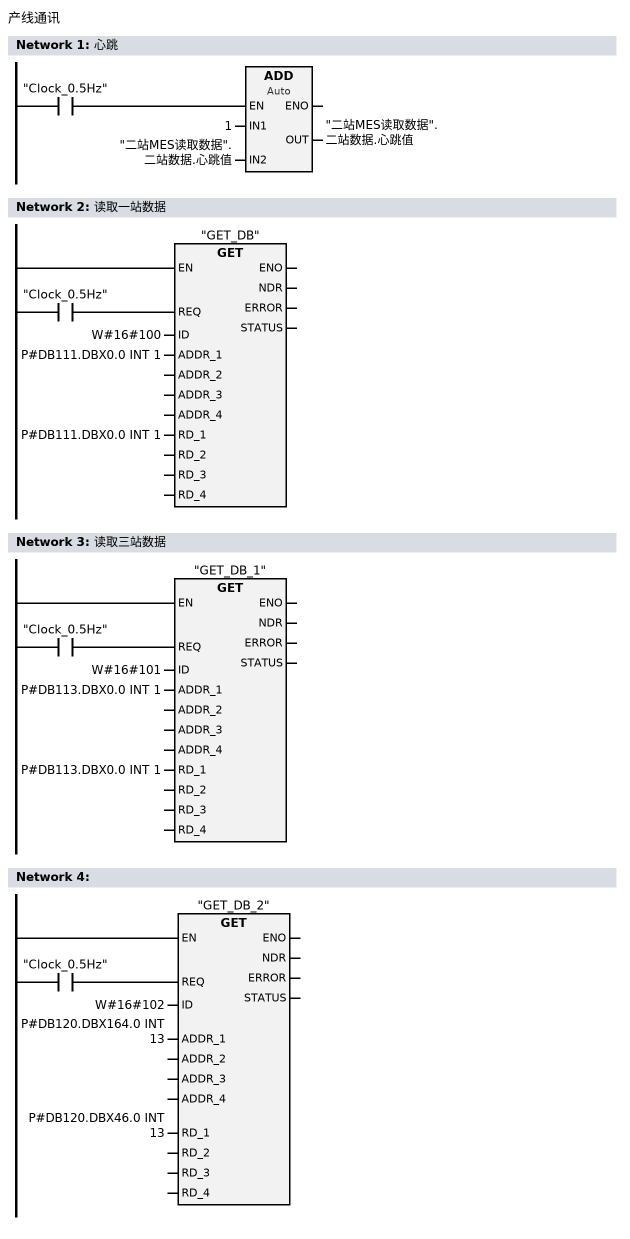
   RUNG wire#powerrail
      Contact( "Clock_0.5Hz" )
      Add(in1 := 1, in2 := "二站MES读取数据".二站数据.心跳值, out => "二站MES读取数据".二站数据.心跳值)
   END_RUNG
   // the same network as SCL:
   IF "Clock_0.5Hz" THEN "二站MES读取数据".二站数据.心跳值 := 1 + "二站MES读取数据".二站数据.心跳值; END_IF;
END_REGION

REGION Network 2: 读取一站数据
   "GET_DB"(REQ := "Clock_0.5Hz", ID := W#16#100, ADDR_1 := P#DB111.DBX0.0 INT 1, RD_1 := P#DB111.DBX0.0 INT 1);   // GET
END_REGION

REGION Network 3: 读取三站数据
   "GET_DB_1"(REQ := "Clock_0.5Hz",   // GET
              ID := W#16#101,
              ADDR_1 := P#DB113.DBX0.0 INT 1,
              RD_1 := P#DB113.DBX0.0 INT 1);
END_REGION

REGION Network 4
   "GET_DB_2"(REQ := "Clock_0.5Hz",   // GET
              ID := W#16#102,
              ADDR_1 := P#DB120.DBX164.0 INT 13,
              RD_1 := P#DB120.DBX46.0 INT 13);
END_REGION
END_FUNCTION

FUNCTION "扫码器通讯" : Void   // FC8, LAD
{ S7_Optimized_Access := 'TRUE' }
VERSION : 0.1
BEGIN

REGION Network 1
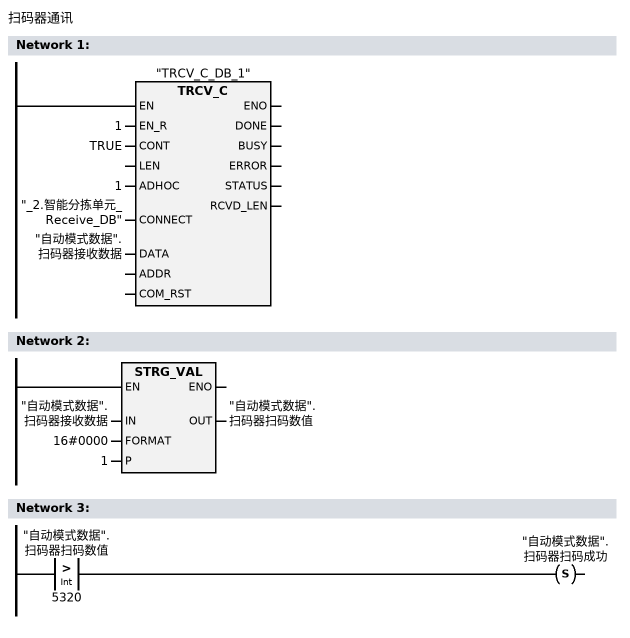
   "TRCV_C_DB_1"(EN_R := 1,   // TRCV_C
                 CONT := TRUE,
                 ADHOC := 1,
                 CONNECT := "_2.智能分拣单元_Receive_DB",
                 DATA := "自动模式数据".扫码器接收数据);
END_REGION

REGION Network 2
   STRG_VAL(IN := "自动模式数据".扫码器接收数据, FORMAT := 16#0000, P := 1, OUT => "自动模式数据".扫码器扫码数值);
END_REGION

REGION Network 3
   RUNG wire#powerrail
      { S7_Templates := "SrcType := Int" } GT_Contact(in1 := "自动模式数据".扫码器扫码数值, in2 := 5320)
      S_Coil( "自动模式数据".扫码器扫码成功 )
   END_RUNG
   // the same network as SCL:
   IF "自动模式数据".扫码器扫码数值 > 5320 THEN "自动模式数据".扫码器扫码成功 := TRUE; END_IF;
END_REGION
END_FUNCTION

FUNCTION "虚拟联动映射" : Void   // FC11, LAD
{ S7_Optimized_Access := 'TRUE' }
VERSION : 0.1
BEGIN

REGION Network 1
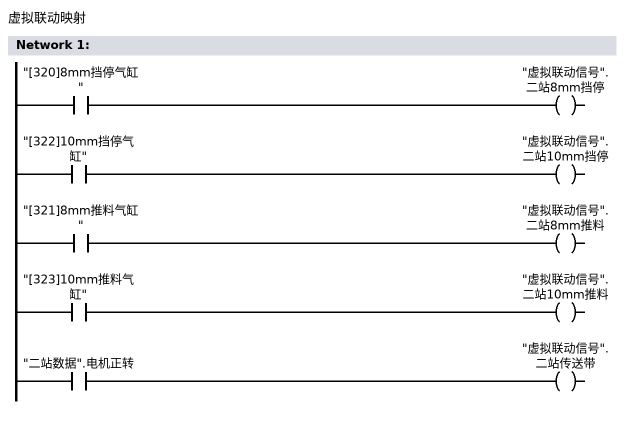
   RUNG wire#powerrail
      Contact( "[320]8mm挡停气缸" )
      Coil( "虚拟联动信号".二站8mm挡停 )
   END_RUNG
   RUNG wire#powerrail
      Contact( "[322]10mm挡停气缸" )
      Coil( "虚拟联动信号".二站10mm挡停 )
   END_RUNG
   RUNG wire#powerrail
      Contact( "[321]8mm推料气缸" )
      Coil( "虚拟联动信号".二站8mm推料 )
   END_RUNG
   RUNG wire#powerrail
      Contact( "[323]10mm推料气缸" )
      Coil( "虚拟联动信号".二站10mm推料 )
   END_RUNG
   RUNG wire#powerrail
      Contact( "二站数据".电机正转 )
      Coil( "虚拟联动信号".二站传送带 )
   END_RUNG
   // the same network as SCL:
   "虚拟联动信号".二站8mm挡停 := "[320]8mm挡停气缸";
   "虚拟联动信号".二站10mm挡停 := "[322]10mm挡停气缸";
   "虚拟联动信号".二站8mm推料 := "[321]8mm推料气缸";
   "虚拟联动信号".二站10mm推料 := "[323]10mm推料气缸";
   "虚拟联动信号".二站传送带 := "二站数据".电机正转;
END_REGION
END_FUNCTION

FUNCTION "AI视觉信号映射" : Void   // FC12, LAD
{ S7_Optimized_Access := 'TRUE' }
VERSION : 0.1
BEGIN

REGION Network 1
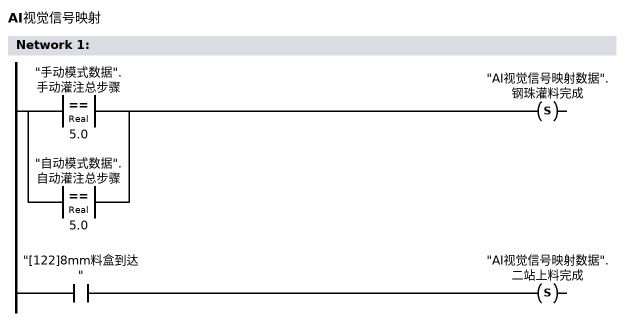
   RUNG wire#powerrail
      { S7_Templates := "SrcType := Real" } EQ_Contact(in1 := "手动模式数据".手动灌注总步骤, in2 := 5.0)
      wire#w1
      S_Coil( "AI视觉信号映射数据".钢珠灌料完成 )
   END_RUNG
   RUNG wire#powerrail
      { S7_Templates := "SrcType := Real" } EQ_Contact(in1 := "自动模式数据".自动灌注总步骤, in2 := 5.0)
   END_RUNG wire#w1
   RUNG wire#powerrail
      Contact( "[122]8mm料盒到达" )
      S_Coil( "AI视觉信号映射数据".二站上料完成 )
   END_RUNG
   // the same network as SCL:
   IF ("手动模式数据".手动灌注总步骤 = 5.0) OR ("自动模式数据".自动灌注总步骤 = 5.0) THEN "AI视觉信号映射数据".钢珠灌料完成 := TRUE; END_IF;
   IF "[122]8mm料盒到达" THEN "AI视觉信号映射数据".二站上料完成 := TRUE; END_IF;
END_REGION
END_FUNCTION

FUNCTION "MES数据映射" : Void   // FC15, LAD
{ S7_Optimized_Access := 'TRUE' }
VERSION : 0.1
BEGIN
END_FUNCTION

// ===== PLC "3.智能仓储单元"  CPU 1214C DC/DC/DC =====

VAR_GLOBAL   // PLC tag table "默认变量表"
   "System_Byte" AT %MB501 : Byte;
   "FirstScan" AT %M501.0 : Bool;
   "DiagStatusUpdate" AT %M501.1 : Bool;
   "AlwaysTRUE" AT %M501.2 : Bool;
   "AlwaysFALSE" AT %M501.3 : Bool;
   "Clock_Byte" AT %MB500 : Byte;
   "Clock_10Hz" AT %M500.0 : Bool;
   "Clock_5Hz" AT %M500.1 : Bool;
   "Clock_2.5Hz" AT %M500.2 : Bool;
   "Clock_2Hz" AT %M500.3 : Bool;
   "Clock_1.25Hz" AT %M500.4 : Bool;
   "Clock_1Hz" AT %M500.5 : Bool;
   "Clock_0.625Hz" AT %M500.6 : Bool;
   "Clock_0.5Hz" AT %M500.7 : Bool;
END_VAR

VAR_GLOBAL   // PLC tag table "第三站变量表"
   "[100]变频编码器" AT %I0.0 : Bool;
   "[101]X伺服左极限" AT %I0.1 : Bool;
   "[102]X伺服右极限" AT %I0.2 : Bool;
   "[103]X伺服原点" AT %I0.3 : Bool;
   "[104]Y伺服左极限" AT %I0.4 : Bool;
   "[105]Y伺服右极限" AT %I0.5 : Bool;
   "[106]Y原点" AT %I0.6 : Bool;
   "[107]启动" AT %I0.7 : Bool;
   "[110]停止" AT %I1.0 : Bool;
   "[111]复位" AT %I1.1 : Bool;
   "[112]急停" AT %I1.2 : Bool;
   "[113]手自动" AT %I1.3 : Bool;
   "[114]盒盖有无检测" AT %I1.4 : Bool;
   "[115]压力检测" AT %I1.5 : Bool;
   "[120]料盒到位检测" AT %I2.0 : Bool;
   "[121]不合格挡料伸出位" AT %I2.1 : Bool;
   "[122]不合格挡料缩回位" AT %I2.2 : Bool;
   "[123]滑台伸出到位" AT %I2.3 : Bool;
   "[124]滑台缩回到位" AT %I2.4 : Bool;
   "[125]]滑台左位" AT %I2.5 : Bool;
   "[126]滑台右位" AT %I2.6 : Bool;
   "[127]滑台夹爪夹紧" AT %I2.7 : Bool;
   "[130]滑台夹爪松开" AT %I3.0 : Bool;
   "[131]不合格推料伸出位" AT %I3.1 : Bool;
   "[132]不合格推料缩回位" AT %I3.2 : Bool;
   "[133]盒盖推料伸出位" AT %I3.3 : Bool;
   "[134]盒盖推料缩回位" AT %I3.4 : Bool;
   "[135]取盒盖伸出位" AT %I3.5 : Bool;
   "[136]取盒盖缩回位" AT %I3.6 : Bool;
   "[137]仓储夹爪夹紧位" AT %I3.7 : Bool;
   "[140]取盒盖上升位" AT %I4.0 : Bool;
   "[141]取盒盖下降位" AT %I4.1 : Bool;
   "[142]仓储伸出位" AT %I4.2 : Bool;
   "[143]仓储缩回位" AT %I4.3 : Bool;
   "[144]仓储上升位" AT %I4.4 : Bool;
   "[145]仓储下降位" AT %I4.5 : Bool;
   "[146]仓储夹爪松开位" AT %I4.6 : Bool;
   "[147]取料挡料伸出位" AT %I4.7 : Bool;
   "[150]取料挡料缩回位" AT %I5.0 : Bool;
   "[151]备用" AT %I5.1 : Bool;
   "[152]备用" AT %I5.2 : Bool;
   "[153]备用" AT %I5.3 : Bool;
   "轴_1_Drive_IN" AT %I68.0 : "PD_TEL3_IN";
   "轴_1_Drive_IN(1)" AT %I86.0 : "PD_TEL3_IN";
   "仓位信息" AT %IW4 : Word;
   "[303]黄色指示灯" AT %Q0.3 : Bool;
   "[304]绿色指示灯" AT %Q0.4 : Bool;
   "[305]红色指示灯" AT %Q0.5 : Bool;
   "[306]变频正转" AT %Q0.6 : Bool;
   "[307]变频反转" AT %Q0.7 : Bool;
   "[310]声光报警" AT %Q1.0 : Bool;
   "[320]不合格挡料气缸" AT %Q2.0 : Bool;
   "[321滑台伸缩气缸" AT %Q2.1 : Bool;
   "[322]滑台移动气缸" AT %Q2.2 : Bool;
   "[323]滑台夹爪气缸" AT %Q2.3 : Bool;
   "[324]不合格推料气缸" AT %Q2.4 : Bool;
   "[325]称重抬升气缸" AT %Q2.5 : Bool;
   "[326]盒盖推料气缸" AT %Q2.6 : Bool;
   "[327]取盖伸缩气缸" AT %Q2.7 : Bool;
   "[330]取盖升降气缸" AT %Q3.0 : Bool;
   "[331]取盖吸盘" AT %Q3.1 : Bool;
   "[332]仓储伸缩气缸" AT %Q3.2 : Bool;
   "[333]仓储升降气缸" AT %Q3.3 : Bool;
   "[334]仓储夹爪控制" AT %Q3.4 : Bool;
   "[335]三色灯-黄" AT %Q3.5 : Bool;
   "[336]三色灯-绿" AT %Q3.6 : Bool;
   "[337]三色灯-红" AT %Q3.7 : Bool;
   "轴_1_Drive_OUT" AT %Q64.0 : "PD_TEL3_OUT";
   "轴_1_Drive_OUT(1)" AT %Q74.0 : "PD_TEL3_OUT";
   "[154]备用4" AT %I5.4 : Bool;
   "[155]变频器故障" AT %I5.5 : Bool;
   "[156]安全光栅" AT %I5.6 : Bool;   // 1无物体2有物体
   "[157]仓位1号有无" AT %I5.7 : Bool;
   "[160]仓位2号有无" AT %I6.0 : Bool;
   "[161]仓位3号有无" AT %I6.1 : Bool;
   "[162]仓位4号有无" AT %I6.2 : Bool;
   "[163]仓位5号有无" AT %I6.3 : Bool;
   "[164]仓位6号有无" AT %I6.4 : Bool;
   "[165]仓位7号有无" AT %I6.5 : Bool;
   "[166]仓位8号有无" AT %I6.6 : Bool;
   "[167]仓位9号有无" AT %I6.7 : Bool;
   "[171]颜色检测" AT %I7.1 : Bool;
   "[170]材质检测" AT %I7.0 : Bool;
   "[311]取料挡料气缸" AT %Q1.1 : Bool;   // 滑台夹爪处挡料气缸
   "[302]备用" AT %I1.6 : Bool;
   "[301]备用" AT %I1.7 : Bool;
   "[300]备用" AT %IW108 : UInt;
   "Tag_4" AT %IW157 : Word;
   "Tag_1" AT %Q0.0 : Bool;
END_VAR

DATA_BLOCK "全局数据块"   // DB5
{ S7_Optimized_Access := 'FALSE' }
VERSION : 0.1
   VAR
      视觉检测步骤 : Real;
      称重压盖步骤 : Real;
      料盒入库步骤 : Real;
      仓储总步骤 : Real;
      重量存储库 : Struct
         "1" : Int;
         "2" : Int;
         "3" : Int;
         "4" : Int;
         "5" : Int;
         "6" : Int;
         "7" : Int;
         "8" : Int;
      END_STRUCT;
      变频器启动 : Bool;
      入站扫码数据 : String[16];
      入站扫码数值 : Int;
      入站扫码成功 : Bool;
      入库扫码数据 : String[16];
      入库扫码数值 : Int;
      入库扫码成功 : Bool;
      视觉检测等待时间 : Time := T#2S;
      不合格产品计数 : Int;
      合格产品计数 : Int;
      上个完成订单ID : Int;
      手动模式步骤 : Real;
      手动存储仓位 : Int := 5;
   END_VAR
BEGIN
END_DATA_BLOCK

DATA_BLOCK "初始化数据"   // DB8
{ S7_Optimized_Access := 'FALSE' }
VERSION : 0.1
   VAR
      手动模式 : Bool;
      自动模式 : Bool;
      自动运行模式 : Bool;
      初始化步骤 : Int;
      初始化完成 : Bool;
      初始化中 : Bool;
      初始化故障 : Bool;
      急停状态 : Bool;
      安全光栅被挡 : Bool;
      黄灯_内部 : Bool;
      红灯_内部 : Bool;
      绿灯_内部 : Bool;
      报警等级 : Int;
      报警确认按钮 : Bool;
      报警总输出 : Bool;
   END_VAR
BEGIN
END_DATA_BLOCK

DATA_BLOCK "状态控制数据"   // DB44
{ S7_Optimized_Access := 'FALSE' }
VERSION : 0.1
   VAR
      在线状态 : Bool;   // PLC已经上电
      忙碌状态 : Bool;   // 三站已经接单
      空闲状态 : Bool;   // 三站准备就绪(没急停，初始化已经完成，光栅没被挡)
      故障状态 : Bool;   // 报警、光栅被挡
   END_VAR
BEGIN
END_DATA_BLOCK

DATA_BLOCK "三站MES读取数据"   // DB120
{ S7_Optimized_Access := 'FALSE' }
VERSION : 0.1
   VAR
      三站数据 : Struct
         在线状态 : Int;
         运行模式 : Int;   // 0 手动 / 1 自动待机 / 2 自动运行
         忙碌状态 : Int;   // 0 空闲 / 1 忙碌
         故障状态 : Int;   // 0 = 无故障
         当前订单ID : Int;   // 当前处理的订单
         当前步骤 : Real;
         心跳值 : Int;
         三站完成 : Bool;
         保留 : Bool;
         保留_1 : Bool;
         保留_2 : Bool;
         保留_3 : Bool;
         保留_4 : Bool;
         保留_5 : Bool;
         保留_6 : Bool;
         仓位状态 : Array[0..8] of Bool;
         入站扫码数据 : Int;
         入库扫码数据 : Int;
         称重数据 : Int;
         产品合格状态 : Int;
         合格产品计数 : Int;
         不合格产品计数 : Int;
         X轴当前位置 : Real;
         Y轴当前位置 : Real;
         完成订单ID : Int;
         三站保留数据 : Array[0..8] of Int;
      END_STRUCT;
      订单数据 : Struct
         订单id : Int;
         ab物料 : Int;   // 1A，2B，3不需要
         小钢珠数量 : Int;
         大钢珠数量 : Int;
         存储仓位 : Int;
         当前订单完成 : Bool;
         开始信号 : Int;
         复位信号 : Int;
         订单保留数据 : Array[0..4] of Int;
      END_STRUCT;
   END_VAR
BEGIN
END_DATA_BLOCK

// folder: System blocks/Program resources

DATA_BLOCK "IEC_Timer_0_DB_7"   // DB7
{ S7_Optimized_Access := 'TRUE' }
AUTHOR : Simatic
FAMILY : IEC
NAME : IEC_TMR
VERSION : 1.0
// stored: InstanceOfName IEC_TIMER
"IEC_TIMER"
BEGIN
END_DATA_BLOCK

DATA_BLOCK "IEC_Timer_0_DB_4"   // DB9
{ S7_Optimized_Access := 'TRUE' }
AUTHOR : Simatic
FAMILY : IEC
NAME : IEC_TMR
VERSION : 1.0
// stored: InstanceOfName IEC_TIMER
"IEC_TIMER"
BEGIN
END_DATA_BLOCK

DATA_BLOCK "IEC_Timer_0_DB"   // DB13
{ S7_Optimized_Access := 'TRUE' }
AUTHOR : Simatic
FAMILY : IEC
NAME : IEC_TMR
VERSION : 1.0
// stored: InstanceOfName IEC_TIMER
"IEC_TIMER"
BEGIN
END_DATA_BLOCK

DATA_BLOCK "IEC_Timer_0_DB_1"   // DB14
{ S7_Optimized_Access := 'TRUE' }
AUTHOR : Simatic
FAMILY : IEC
NAME : IEC_TMR
VERSION : 1.0
// stored: InstanceOfName IEC_TIMER
"IEC_TIMER"
BEGIN
END_DATA_BLOCK

DATA_BLOCK "IEC_Timer_0_DB_2"   // DB15
{ S7_Optimized_Access := 'TRUE' }
AUTHOR : Simatic
FAMILY : IEC
NAME : IEC_TMR
VERSION : 1.0
// stored: InstanceOfName IEC_TIMER
"IEC_TIMER"
BEGIN
END_DATA_BLOCK

DATA_BLOCK "IEC_Timer_0_DB_3"   // DB16
{ S7_Optimized_Access := 'TRUE' }
AUTHOR : Simatic
FAMILY : IEC
NAME : IEC_TMR
VERSION : 1.0
// stored: InstanceOfName IEC_TIMER
"IEC_TIMER"
BEGIN
END_DATA_BLOCK

DATA_BLOCK "IEC_Timer_0_DB_5"   // DB18
{ S7_Optimized_Access := 'TRUE' }
AUTHOR : Simatic
FAMILY : IEC
NAME : IEC_TMR
VERSION : 1.0
// stored: InstanceOfName IEC_TIMER
"IEC_TIMER"
BEGIN
END_DATA_BLOCK

DATA_BLOCK "IEC_Timer_0_DB_6"   // DB19
{ S7_Optimized_Access := 'TRUE' }
AUTHOR : Simatic
FAMILY : IEC
NAME : IEC_TMR
VERSION : 1.0
// stored: InstanceOfName IEC_TIMER
"IEC_TIMER"
BEGIN
END_DATA_BLOCK

DATA_BLOCK "IEC_Timer_0_DB_8"   // DB28
{ S7_Optimized_Access := 'TRUE' }
AUTHOR : Simatic
FAMILY : IEC
NAME : IEC_TMR
VERSION : 1.0
// stored: InstanceOfName IEC_TIMER
"IEC_TIMER"
BEGIN
END_DATA_BLOCK

DATA_BLOCK "IEC_Timer_0_DB_9"   // DB29
{ S7_Optimized_Access := 'TRUE' }
AUTHOR : Simatic
FAMILY : IEC
NAME : IEC_TMR
VERSION : 1.0
// stored: InstanceOfName IEC_TIMER
"IEC_TIMER"
BEGIN
END_DATA_BLOCK

DATA_BLOCK "IEC_Timer_0_DB_10"   // DB30
{ S7_Optimized_Access := 'TRUE' }
AUTHOR : Simatic
FAMILY : IEC
NAME : IEC_TMR
VERSION : 1.0
// stored: InstanceOfName IEC_TIMER
"IEC_TIMER"
BEGIN
END_DATA_BLOCK

DATA_BLOCK "IEC_Timer_0_DB_11"   // DB31
{ S7_Optimized_Access := 'TRUE' }
AUTHOR : Simatic
FAMILY : IEC
NAME : IEC_TMR
VERSION : 1.0
// stored: InstanceOfName IEC_TIMER
"IEC_TIMER"
BEGIN
END_DATA_BLOCK

DATA_BLOCK "IEC_Timer_0_DB_12"   // DB32
{ S7_Optimized_Access := 'TRUE' }
AUTHOR : Simatic
FAMILY : IEC
NAME : IEC_TMR
VERSION : 1.0
// stored: InstanceOfName IEC_TIMER
"IEC_TIMER"
BEGIN
END_DATA_BLOCK

DATA_BLOCK "IEC_Timer_0_DB_13"   // DB33
{ S7_Optimized_Access := 'TRUE' }
AUTHOR : Simatic
FAMILY : IEC
NAME : IEC_TMR
VERSION : 1.0
// stored: InstanceOfName IEC_TIMER
"IEC_TIMER"
BEGIN
END_DATA_BLOCK

DATA_BLOCK "_3.智能仓储单元_Receive_DB"   // DB35
{ S7_Optimized_Access := 'TRUE' }
AUTHOR : SIMATIC
FAMILY : MC7Plus
NAME : TC_IP_v4
VERSION : 1.0
// stored: InstanceOfName TCON_IP_v4
"TCON_IP_v4"
BEGIN
   ID := 104;
   InterfaceId := 64;
   LocalPort := 8899;
   RemotePort := 8899;
   RemoteAddress.ADDR[1] := 192;
   RemoteAddress.ADDR[2] := 168;
   RemoteAddress.ADDR[3] := 40;
   RemoteAddress.ADDR[4] := 103;
END_DATA_BLOCK

DATA_BLOCK "IEC_Timer_0_DB_17"   // DB37
{ S7_Optimized_Access := 'TRUE' }
AUTHOR : Simatic
FAMILY : IEC
NAME : IEC_TMR
VERSION : 1.0
// stored: InstanceOfName IEC_TIMER
"IEC_TIMER"
BEGIN
END_DATA_BLOCK

DATA_BLOCK "IEC_Timer_0_DB_18"   // DB38
{ S7_Optimized_Access := 'TRUE' }
AUTHOR : Simatic
FAMILY : IEC
NAME : IEC_TMR
VERSION : 1.0
// stored: InstanceOfName IEC_TIMER
"IEC_TIMER"
BEGIN
END_DATA_BLOCK

DATA_BLOCK "IEC_Timer_0_DB_19"   // DB39
{ S7_Optimized_Access := 'TRUE' }
AUTHOR : Simatic
FAMILY : IEC
NAME : IEC_TMR
VERSION : 1.0
// stored: InstanceOfName IEC_TIMER
"IEC_TIMER"
BEGIN
END_DATA_BLOCK

DATA_BLOCK "IEC_Timer_0_DB_16"   // DB40
{ S7_Optimized_Access := 'TRUE' }
AUTHOR : Simatic
FAMILY : IEC
NAME : IEC_TMR
VERSION : 1.0
// stored: InstanceOfName IEC_TIMER
"IEC_TIMER"
BEGIN
END_DATA_BLOCK

DATA_BLOCK "_3.智能仓储单元_Receive_DB_1"   // DB41
{ S7_Optimized_Access := 'TRUE' }
AUTHOR : SIMATIC
FAMILY : MC7Plus
NAME : TC_IP_v4
VERSION : 1.0
// stored: InstanceOfName TCON_IP_v4
"TCON_IP_v4"
BEGIN
   ID := 107;
   InterfaceId := 64;
   LocalPort := 8899;
   RemotePort := 8899;
   RemoteAddress.ADDR[1] := 192;
   RemoteAddress.ADDR[2] := 168;
   RemoteAddress.ADDR[3] := 40;
   RemoteAddress.ADDR[4] := 102;
END_DATA_BLOCK

DATA_BLOCK "IEC_Timer_0_DB_20"   // DB42
{ S7_Optimized_Access := 'TRUE' }
AUTHOR : Simatic
FAMILY : IEC
NAME : IEC_TMR
VERSION : 1.0
// stored: InstanceOfName IEC_TIMER
"IEC_TIMER"
BEGIN
END_DATA_BLOCK

DATA_BLOCK "IEC_Timer_0_DB_14"   // DB45
{ S7_Optimized_Access := 'TRUE' }
AUTHOR : Simatic
FAMILY : IEC
NAME : IEC_TMR
VERSION : 1.0
// stored: InstanceOfName IEC_TIMER
"IEC_TIMER"
BEGIN
END_DATA_BLOCK

DATA_BLOCK "IEC_Timer_0_DB_15"   // DB46
{ S7_Optimized_Access := 'TRUE' }
AUTHOR : Simatic
FAMILY : IEC
NAME : IEC_TMR
VERSION : 1.0
// stored: InstanceOfName IEC_TIMER
"IEC_TIMER"
BEGIN
END_DATA_BLOCK

DATA_BLOCK "IEC_Timer_0_DB_21"   // DB47
{ S7_Optimized_Access := 'TRUE' }
AUTHOR : Simatic
FAMILY : IEC
NAME : IEC_TMR
VERSION : 1.0
// stored: InstanceOfName IEC_TIMER
"IEC_TIMER"
BEGIN
END_DATA_BLOCK

DATA_BLOCK "IEC_Timer_0_DB_22"   // DB48
{ S7_Optimized_Access := 'TRUE' }
AUTHOR : Simatic
FAMILY : IEC
NAME : IEC_TMR
VERSION : 1.0
// stored: InstanceOfName IEC_TIMER
"IEC_TIMER"
BEGIN
END_DATA_BLOCK

DATA_BLOCK "IEC_Timer_0_DB_23"   // DB49
{ S7_Optimized_Access := 'TRUE' }
AUTHOR : Simatic
FAMILY : IEC
NAME : IEC_TMR
VERSION : 1.0
// stored: InstanceOfName IEC_TIMER
"IEC_TIMER"
BEGIN
END_DATA_BLOCK

DATA_BLOCK "IEC_Timer_0_DB_24"   // DB50
{ S7_Optimized_Access := 'TRUE' }
AUTHOR : Simatic
FAMILY : IEC
NAME : IEC_TMR
VERSION : 1.0
// stored: InstanceOfName IEC_TIMER
"IEC_TIMER"
BEGIN
END_DATA_BLOCK

DATA_BLOCK "IEC_Timer_0_DB_25"   // DB51
{ S7_Optimized_Access := 'TRUE' }
AUTHOR : Simatic
FAMILY : IEC
NAME : IEC_TMR
VERSION : 1.0
// stored: InstanceOfName IEC_TIMER
"IEC_TIMER"
BEGIN
END_DATA_BLOCK

DATA_BLOCK "IEC_Timer_0_DB_26"   // DB52
{ S7_Optimized_Access := 'TRUE' }
AUTHOR : Simatic
FAMILY : IEC
NAME : IEC_TMR
VERSION : 1.0
// stored: InstanceOfName IEC_TIMER
"IEC_TIMER"
BEGIN
END_DATA_BLOCK

DATA_BLOCK "IEC_Timer_0_DB_27"   // DB53
{ S7_Optimized_Access := 'TRUE' }
AUTHOR : Simatic
FAMILY : IEC
NAME : IEC_TMR
VERSION : 1.0
// stored: InstanceOfName IEC_TIMER
"IEC_TIMER"
BEGIN
END_DATA_BLOCK

DATA_BLOCK "IEC_Timer_0_DB_28"   // DB54
{ S7_Optimized_Access := 'TRUE' }
AUTHOR : Simatic
FAMILY : IEC
NAME : IEC_TMR
VERSION : 1.0
// stored: InstanceOfName IEC_TIMER
"IEC_TIMER"
BEGIN
END_DATA_BLOCK

DATA_BLOCK "IEC_Timer_0_DB_29"   // DB55
{ S7_Optimized_Access := 'TRUE' }
AUTHOR : Simatic
FAMILY : IEC
NAME : IEC_TMR
VERSION : 1.0
// stored: InstanceOfName IEC_TIMER
"IEC_TIMER"
BEGIN
END_DATA_BLOCK

DATA_BLOCK "IEC_Timer_0_DB_30"   // DB56
{ S7_Optimized_Access := 'TRUE' }
AUTHOR : Simatic
FAMILY : IEC
NAME : IEC_TMR
VERSION : 1.0
// stored: InstanceOfName IEC_TIMER
"IEC_TIMER"
BEGIN
END_DATA_BLOCK

DATA_BLOCK "IEC_Timer_0_DB_31"   // DB57
{ S7_Optimized_Access := 'TRUE' }
AUTHOR : Simatic
FAMILY : IEC
NAME : IEC_TMR
VERSION : 1.0
// stored: InstanceOfName IEC_TIMER
"IEC_TIMER"
BEGIN
END_DATA_BLOCK

DATA_BLOCK "IEC_Timer_0_DB_32"   // DB58
{ S7_Optimized_Access := 'TRUE' }
AUTHOR : Simatic
FAMILY : IEC
NAME : IEC_TMR
VERSION : 1.0
// stored: InstanceOfName IEC_TIMER
"IEC_TIMER"
BEGIN
END_DATA_BLOCK

DATA_BLOCK "IEC_Timer_0_DB_33"   // DB59
{ S7_Optimized_Access := 'TRUE' }
AUTHOR : Simatic
FAMILY : IEC
NAME : IEC_TMR
VERSION : 1.0
// stored: InstanceOfName IEC_TIMER
"IEC_TIMER"
BEGIN
END_DATA_BLOCK

DATA_BLOCK "IEC_Timer_0_DB_34"   // DB60
{ S7_Optimized_Access := 'TRUE' }
AUTHOR : Simatic
FAMILY : IEC
NAME : IEC_TMR
VERSION : 1.0
// stored: InstanceOfName IEC_TIMER
"IEC_TIMER"
BEGIN
END_DATA_BLOCK

DATA_BLOCK "IEC_Timer_0_DB_35"   // DB61
{ S7_Optimized_Access := 'TRUE' }
AUTHOR : Simatic
FAMILY : IEC
NAME : IEC_TMR
VERSION : 1.0
// stored: InstanceOfName IEC_TIMER
"IEC_TIMER"
BEGIN
END_DATA_BLOCK

// folder: 运动控制

DATA_BLOCK "运动控制数据2"   // DB1
{ S7_Optimized_Access := 'FALSE' }
VERSION : 0.1
   VAR
      X轴位置 : Real;
      Y轴位置 : Real;
      称重抓取x值 : Real := -82.0;
      称重抓取y值 : Real := 537.0;
      扫码位x值 : Real := -29.0;
      扫码位y值 : Real := 382.0;
      abc位x值 : Real := 151.0;
      def位x值 : Real := -32.0;
      ghi位x值 : Real := -208.0;
      adg位y值 : Real := -231.0;
      bef位y值 : Real := -51.0;
      cfi位y值 : Real := 121.0;
      "出仓位x值-420.38" : Real := -416.0;
      "出仓位y值162.88" : Real := 152.0;
      X值统一入库位 : Bool;
      Y值统一入库位 : Bool;
      X值计算 : Int;
      Y值计算 : Int;
      Y值转换后 : Int;
   END_VAR
BEGIN
END_DATA_BLOCK

DATA_BLOCK "运动控制数据1"   // DB43
{ S7_Optimized_Access := 'FALSE' }
VERSION : 0.1
   VAR
      轴初始化按钮 : Bool;
      轴初始化完成 : Bool;
      轴初始化步骤 : Int;
      轴初始化错误 : Bool;
      X轴机械手错误输出 : Bool;
      Y轴机械手错误输出 : Bool;
      X轴使能按钮 : Bool;
      X轴使能状态 : Bool;
      X轴使能错误 : Bool;
      X轴复位按钮 : Bool;
      X轴复位完成 : Bool;
      X轴复位错误 : Bool;
      X轴回原位按钮 : Bool;
      X轴回原位完成 : Bool;
      X轴回原位错误 : Bool;
      X轴绝对定位按钮 : Bool;
      X轴绝对定位完成 : Bool;
      X轴绝对定位错误 : Bool;
      Y轴使能按钮 : Bool;
      Y轴使能状态 : Bool;
      Y轴使能错误 : Bool;
      Y轴复位按钮 : Bool;
      Y轴复位完成 : Bool;
      Y轴复位错误 : Bool;
      Y轴回原位按钮 : Bool;
      Y轴回原位完成 : Bool;
      Y轴回原位错误 : Bool;
      Y轴绝对定位按钮 : Bool;
      Y轴绝对定位完成 : Bool;
      Y轴绝对定位错误 : Bool;
   END_VAR
BEGIN
END_DATA_BLOCK

// folder: 通讯模块

DATA_BLOCK "虚实联动信号"   // DB4
{ S7_Optimized_Access := 'FALSE' }
VERSION : 0.1
   VAR
      变频正转 : Bool;
      变频反转 : Bool;
      滑台移动气缸 : Bool;
      滑台伸缩气缸 : Bool;
      仓储伸缩气缸 : Bool;
      仓储升降气缸 : Bool;
      称重抬升气缸 : Bool;
      不合格推料气缸 : Bool;
      不合格挡料气缸 : Bool;
      取料挡料气缸 : Bool;
      取盖伸缩气缸 : Bool;
      取盖升降气缸 : Bool;
      盒盖推料气缸 : Bool;
      滑台夹爪气缸 : Bool;
      仓储夹爪控制 : Bool;
      取盖吸盘 : Bool;
   END_VAR
BEGIN
END_DATA_BLOCK

DATA_BLOCK "称重数据"   // DB12
{ S7_Optimized_Access := 'FALSE' }
VERSION : 0.1
   VAR
      称重 : Struct
         称重数据 : Int;
         称重数据接收 : Int;
      END_STRUCT;
   END_VAR
BEGIN
END_DATA_BLOCK

DATA_BLOCK "一站数据"   // DB111
{ S7_Optimized_Access := 'FALSE' }
VERSION : 0.1
   VAR
      一站完成 : Bool;
      复位完成 : Bool;
      一站就绪 : Bool;
      一站忙碌 : Bool;
      一站请求二站接收 : Bool;
      一站可接单 : Bool;
      数据7 : Bool;
      数据8 : Bool;
      数据9 : Bool;
      数据10 : Bool;
      数据11 : Bool;
      数据12 : Bool;
      数据13 : Bool;
      数据14 : Bool;
   END_VAR
BEGIN
END_DATA_BLOCK

DATA_BLOCK "二站数据"   // DB112
{ S7_Optimized_Access := 'FALSE' }
VERSION : 0.1
   VAR
      二站完成 : Bool;
      二站已接收 : Bool;
      复位完成 : Bool;
      空闲状态 : Bool;
      电机正转 : Bool;
      二站忙碌 : Bool;
      二站请求三站接收 : Bool;
      二站可接收 : Bool;
      数据17 : Bool;
      数据18 : Bool;
      数据19 : Bool;
      数据20 : Bool;
      数据21 : Bool;
   END_VAR
BEGIN
END_DATA_BLOCK

DATA_BLOCK "三站数据"   // DB113
{ S7_Optimized_Access := 'FALSE' }
VERSION : 0.1
   VAR
      三站完成 : Bool;
      三站已接收 : Bool;
      复位完成 : Bool;
      空闲状态 : Bool;
      出现废料 : Bool;
      安全光栅 : Bool;
      三站可接收 : Bool;
      三站忙碌 : Bool;
      数据23 : Bool;
      数据24 : Bool;
      数据25 : Bool;
      数据26 : Bool;
      数据27 : Bool;
      数据28 : Bool;
      数据29 : Bool;
   END_VAR
BEGIN
END_DATA_BLOCK

DATA_BLOCK "AI视觉信号映射数据"   // DB116
{ S7_Optimized_Access := 'TRUE' }
VERSION : 0.1
   VAR
      三站压盖完成 : Bool;
      三站入库完成 : Bool;
   END_VAR
BEGIN
END_DATA_BLOCK

// folder: (top level)

DATA_BLOCK "X轴机械手"   // DB2, Motion_DB
{ S7_Optimized_Access := 'TRUE' }
AUTHOR : SIMATIC
FAMILY : BasicMC
NAME : TO_PosAx
VERSION : 7.0
// stored: InstanceOfName TO_PositioningAxis
"TO_PositioningAxis"
BEGIN
   // Axis.HomingReferencePointSwitch_AddressCU = %I0.3
   // Axis.PositionLimitsMax_AddressCU = %I0.1
   // Axis.PositionLimitsMin_AddressCU = %I0.2
   // Axis.Encoder.TelegramAddressOutCU = %Q74.0
   // Axis.Encoder.TelegramAddressInCU = %I86.0
   // Axis.Encoder.DoNameCU = SINAMICS-V90-PN_2.驱动_1_编码器1
   // Axis.Drive.TelegramAddressOutCU = %Q74.0
   // Axis.Drive.TelegramAddressInCU = %I86.0
   // Axis.Drive.TelegramType = 2
   // Axis.Drive.DoNameCU = SINAMICS-V90-PN_2.驱动_1
   // Axis.LengthUnitNormalized.Distance = 1013
   // Axis.Encoder.SelectedHscIndexCU = -1
   // Axis.Encoder.DbTypeCU = Classic
   // Axis.Drive.DbTypeCU = Classic
END_DATA_BLOCK

DATA_BLOCK "Y轴机械手"   // DB3, Motion_DB
{ S7_Optimized_Access := 'TRUE' }
AUTHOR : SIMATIC
FAMILY : BasicMC
NAME : TO_PosAx
VERSION : 7.0
// stored: InstanceOfName TO_PositioningAxis
"TO_PositioningAxis"
BEGIN
   // Axis.HomingReferencePointSwitch_AddressCU = %I0.6
   // Axis.PositionLimitsMax_AddressCU = %I0.4
   // Axis.PositionLimitsMin_AddressCU = %I0.5
   // Axis.Encoder.TelegramAddressOutCU = %Q64.0
   // Axis.Encoder.TelegramAddressInCU = %I68.0
   // Axis.Encoder.DoNameCU = SINAMICS-V90-PN_1.驱动_1_编码器1
   // Axis.Drive.TelegramAddressOutCU = %Q64.0
   // Axis.Drive.TelegramAddressInCU = %I68.0
   // Axis.Drive.TelegramType = 2
   // Axis.Drive.DoNameCU = SINAMICS-V90-PN_1.驱动_1
   // Axis.LengthUnitNormalized.Distance = 1013
   // Axis.Encoder.SelectedHscIndexCU = -1
   // Axis.Encoder.DbTypeCU = Classic
   // Axis.Drive.DbTypeCU = Classic
END_DATA_BLOCK

FUNCTION "0.初始化" : Void   // FC5, LAD
{ S7_Optimized_Access := 'TRUE' }
VERSION : 0.1
   VAR_TEMP   // added for the SCL form of the ladder/FBD networks
      _w1 : Bool;
      _w2 : Bool;
   END_VAR
BEGIN

REGION Network 1: 模式切换
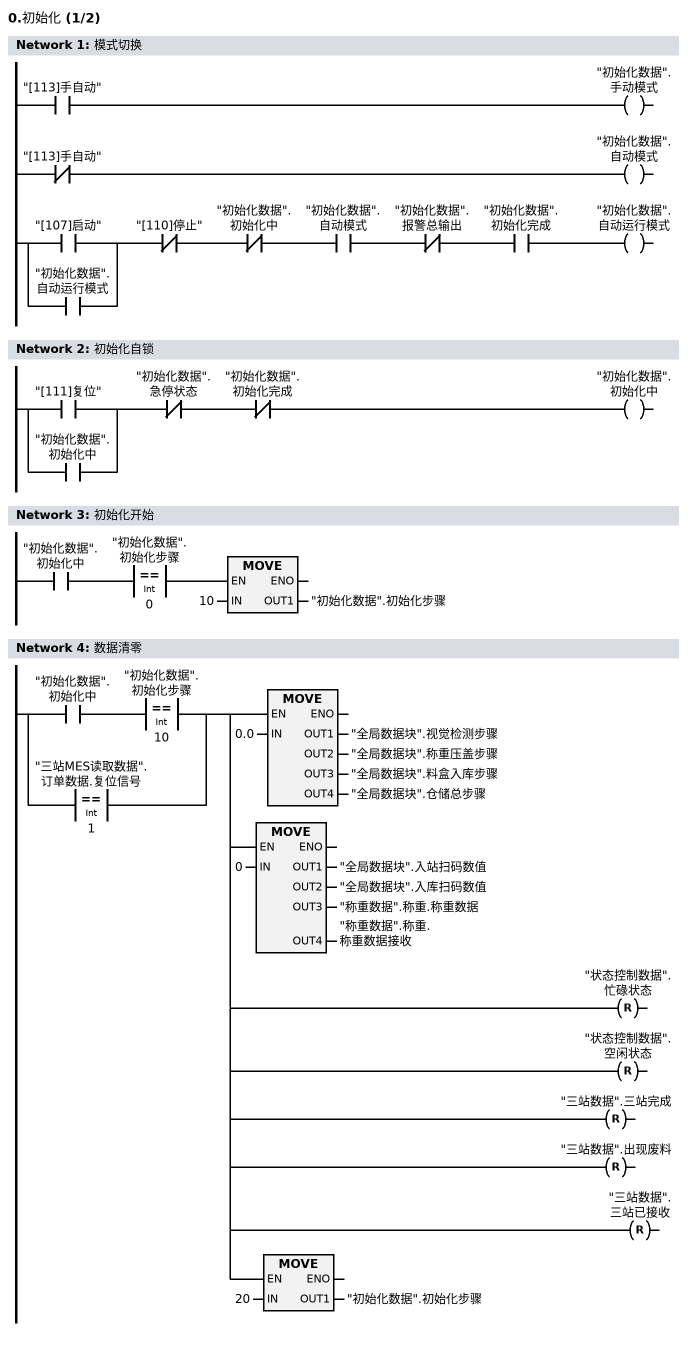
   RUNG wire#powerrail
      Contact( "[113]手自动" )
      Coil( "初始化数据".手动模式 )
   END_RUNG
   RUNG wire#powerrail
      I_Contact( "[113]手自动" )
      Coil( "初始化数据".自动模式 )
   END_RUNG
   RUNG wire#powerrail
      Contact( "[107]启动" )
      wire#w1
      I_Contact( "[110]停止" )
      I_Contact( "初始化数据".初始化中 )
      Contact( "初始化数据".自动模式 )
      I_Contact( "初始化数据".报警总输出 )
      Contact( "初始化数据".初始化完成 )
      Coil( "初始化数据".自动运行模式 )
   END_RUNG
   RUNG wire#powerrail
      Contact( "初始化数据".自动运行模式 )
   END_RUNG wire#w1
   // the same network as SCL:
   "初始化数据".手动模式 := "[113]手自动";
   "初始化数据".自动模式 := NOT "[113]手自动";
   "初始化数据".自动运行模式 := ("[107]启动" OR "初始化数据".自动运行模式) AND NOT "[110]停止" AND NOT "初始化数据".初始化中 AND "初始化数据".自动模式 AND NOT "初始化数据".报警总输出 AND "初始化数据".初始化完成;
END_REGION

REGION Network 2: 初始化自锁
   RUNG wire#powerrail
      Contact( "[111]复位" )
      wire#w1
      I_Contact( "初始化数据".急停状态 )
      I_Contact( "初始化数据".初始化完成 )
      Coil( "初始化数据".初始化中 )
   END_RUNG
   RUNG wire#powerrail
      Contact( "初始化数据".初始化中 )
   END_RUNG wire#w1
   // the same network as SCL:
   "初始化数据".初始化中 := ("[111]复位" OR "初始化数据".初始化中) AND NOT "初始化数据".急停状态 AND NOT "初始化数据".初始化完成;
END_REGION

REGION Network 3: 初始化开始
   RUNG wire#powerrail
      Contact( "初始化数据".初始化中 )
      { S7_Templates := "SrcType := Int" } EQ_Contact(in1 := "初始化数据".初始化步骤, in2 := 0)
      Move(in := 10, out1 => "初始化数据".初始化步骤)
   END_RUNG
   // the same network as SCL:
   IF "初始化数据".初始化中 AND ("初始化数据".初始化步骤 = 0) THEN "初始化数据".初始化步骤 := 10; END_IF;
END_REGION

REGION Network 4: 数据清零
   RUNG wire#powerrail
      Contact( "初始化数据".初始化中 )
      { S7_Templates := "SrcType := Int" } EQ_Contact(in1 := "初始化数据".初始化步骤, in2 := 10)
      wire#w1
      Move(in := 0.0, out1 => "全局数据块".视觉检测步骤, out2 => "全局数据块".称重压盖步骤, out3 => "全局数据块".料盒入库步骤, out4 => "全局数据块".仓储总步骤)
   END_RUNG
   RUNG wire#powerrail
      { S7_Templates := "SrcType := Int" } EQ_Contact(in1 := "三站MES读取数据".订单数据.复位信号, in2 := 1)
   END_RUNG wire#w1
   RUNG wire#w1
      Move(in := 0, out1 => "全局数据块".入站扫码数值, out2 => "全局数据块".入库扫码数值, out3 => "称重数据".称重.称重数据, out4 => "称重数据".称重.称重数据接收)
   END_RUNG
   RUNG wire#w1
      R_Coil( "状态控制数据".忙碌状态 )
   END_RUNG
   RUNG wire#w1
      R_Coil( "状态控制数据".空闲状态 )
   END_RUNG
   RUNG wire#w1
      R_Coil( "三站数据".三站完成 )
   END_RUNG
   RUNG wire#w1
      R_Coil( "三站数据".出现废料 )
   END_RUNG
   RUNG wire#w1
      R_Coil( "三站数据".三站已接收 )
   END_RUNG
   RUNG wire#w1
      Move(in := 20, out1 => "初始化数据".初始化步骤)
   END_RUNG
   // the same network as SCL:
   IF ("初始化数据".初始化中 AND ("初始化数据".初始化步骤 = 10)) OR ("三站MES读取数据".订单数据.复位信号 = 1) THEN
       "全局数据块".视觉检测步骤 := 0.0;
       "全局数据块".称重压盖步骤 := 0.0;
       "全局数据块".料盒入库步骤 := 0.0;
       "全局数据块".仓储总步骤 := 0.0;
       "全局数据块".入站扫码数值 := 0;
       "全局数据块".入库扫码数值 := 0;
       "称重数据".称重.称重数据 := 0;
       "称重数据".称重.称重数据接收 := 0;
       "状态控制数据".忙碌状态 := FALSE;
       "状态控制数据".空闲状态 := FALSE;
       "三站数据".三站完成 := FALSE;
       "三站数据".出现废料 := FALSE;
       "三站数据".三站已接收 := FALSE;
       "初始化数据".初始化步骤 := 20;
   END_IF;
END_REGION

REGION Network 6: 气缸复位
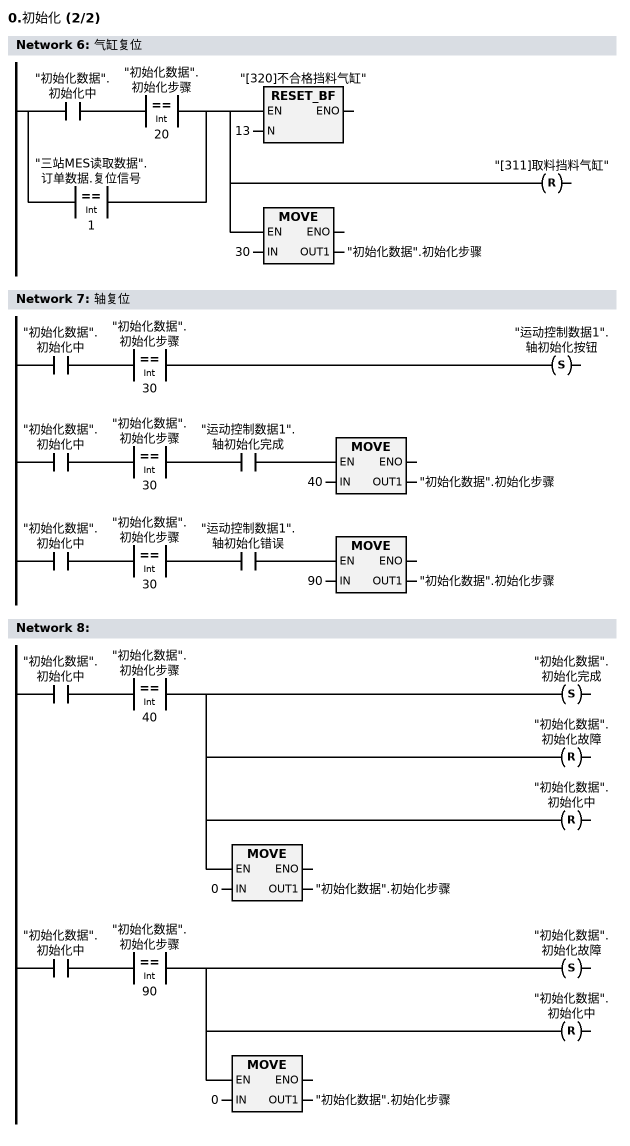
   // no SCL statement known for RBitfield: written as a call
   #_w1 := ("初始化数据".初始化中 AND ("初始化数据".初始化步骤 = 20)) OR ("三站MES读取数据".订单数据.复位信号 = 1);
   IF #_w1 THEN
       RESET_BF(operand := "[320]不合格挡料气缸", n := 13);
       "[311]取料挡料气缸" := FALSE;
       "初始化数据".初始化步骤 := 30;
   END_IF;
END_REGION

REGION Network 7: 轴复位
   RUNG wire#powerrail
      Contact( "初始化数据".初始化中 )
      { S7_Templates := "SrcType := Int" } EQ_Contact(in1 := "初始化数据".初始化步骤, in2 := 30)
      S_Coil( "运动控制数据1".轴初始化按钮 )
   END_RUNG
   RUNG wire#powerrail
      Contact( "初始化数据".初始化中 )
      { S7_Templates := "SrcType := Int" } EQ_Contact(in1 := "初始化数据".初始化步骤, in2 := 30)
      Contact( "运动控制数据1".轴初始化完成 )
      Move(in := 40, out1 => "初始化数据".初始化步骤)
   END_RUNG
   RUNG wire#powerrail
      Contact( "初始化数据".初始化中 )
      { S7_Templates := "SrcType := Int" } EQ_Contact(in1 := "初始化数据".初始化步骤, in2 := 30)
      Contact( "运动控制数据1".轴初始化错误 )
      Move(in := 90, out1 => "初始化数据".初始化步骤)
   END_RUNG
   // the same network as SCL:
   IF "初始化数据".初始化中 AND ("初始化数据".初始化步骤 = 30) THEN "运动控制数据1".轴初始化按钮 := TRUE; END_IF;
   IF "初始化数据".初始化中 AND ("初始化数据".初始化步骤 = 30) AND "运动控制数据1".轴初始化完成 THEN "初始化数据".初始化步骤 := 40; END_IF;
   IF "初始化数据".初始化中 AND ("初始化数据".初始化步骤 = 30) AND "运动控制数据1".轴初始化错误 THEN "初始化数据".初始化步骤 := 90; END_IF;
END_REGION

REGION Network 8
   RUNG wire#powerrail
      Contact( "初始化数据".初始化中 )
      { S7_Templates := "SrcType := Int" } EQ_Contact(in1 := "初始化数据".初始化步骤, in2 := 40)
      wire#w1
      S_Coil( "初始化数据".初始化完成 )
   END_RUNG
   RUNG wire#w1
      R_Coil( "初始化数据".初始化故障 )
   END_RUNG
   RUNG wire#w1
      R_Coil( "初始化数据".初始化中 )
   END_RUNG
   RUNG wire#w1
      Move(in := 0, out1 => "初始化数据".初始化步骤)
   END_RUNG
   RUNG wire#powerrail
      Contact( "初始化数据".初始化中 )
      { S7_Templates := "SrcType := Int" } EQ_Contact(in1 := "初始化数据".初始化步骤, in2 := 90)
      wire#w2
      S_Coil( "初始化数据".初始化故障 )
   END_RUNG
   RUNG wire#w2
      R_Coil( "初始化数据".初始化中 )
   END_RUNG
   RUNG wire#w2
      Move(in := 0, out1 => "初始化数据".初始化步骤)
   END_RUNG
   // the same network as SCL:
   IF "初始化数据".初始化中 AND ("初始化数据".初始化步骤 = 40) THEN
       "初始化数据".初始化完成 := TRUE;
       "初始化数据".初始化故障 := FALSE;
   END_IF;
   #_w1 := "初始化数据".初始化中 AND ("初始化数据".初始化步骤 = 40);
   IF #_w1 THEN
       "初始化数据".初始化中 := FALSE;
       "初始化数据".初始化步骤 := 0;
   END_IF;
   IF "初始化数据".初始化中 AND ("初始化数据".初始化步骤 = 90) THEN "初始化数据".初始化故障 := TRUE; END_IF;
   #_w2 := "初始化数据".初始化中 AND ("初始化数据".初始化步骤 = 90);
   IF #_w2 THEN
       "初始化数据".初始化中 := FALSE;
       "初始化数据".初始化步骤 := 0;
   END_IF;
END_REGION
END_FUNCTION

FUNCTION "2.状态控制" : Void   // FC6, LAD
{ S7_Optimized_Access := 'TRUE' }
VERSION : 0.1
BEGIN

REGION Network 1: 三站四种状态
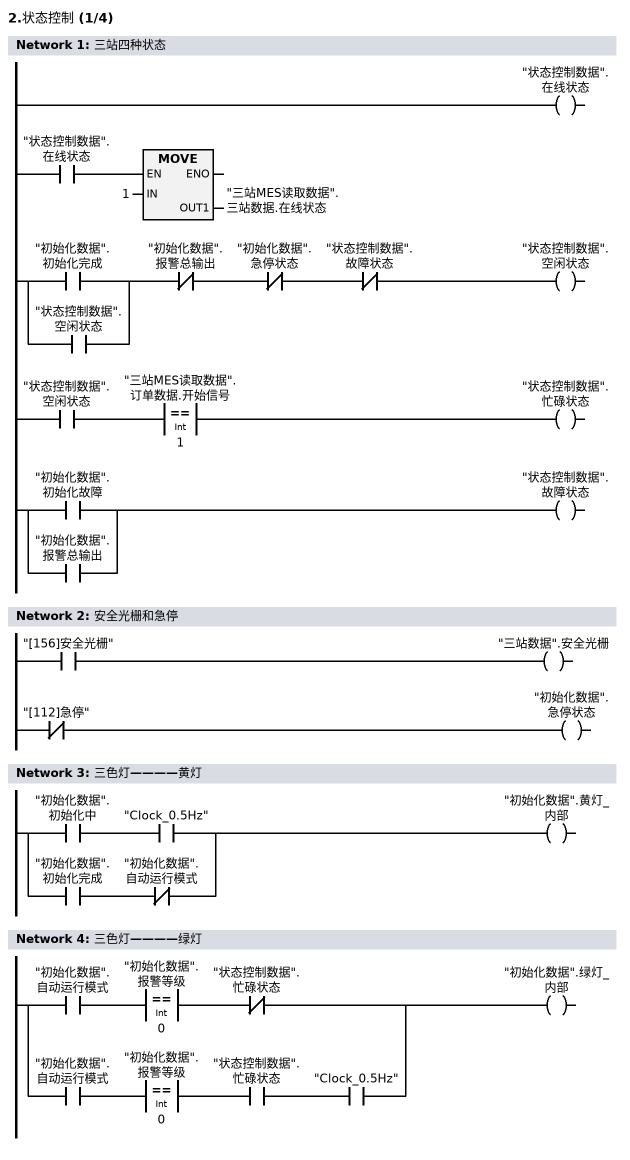
   RUNG wire#powerrail
      Coil( "状态控制数据".在线状态 )
   END_RUNG
   RUNG wire#powerrail
      Contact( "状态控制数据".在线状态 )
      Move(in := 1, out1 => "三站MES读取数据".三站数据.在线状态)
   END_RUNG
   RUNG wire#powerrail
      Contact( "初始化数据".初始化完成 )
      wire#w1
      I_Contact( "初始化数据".报警总输出 )
      I_Contact( "初始化数据".急停状态 )
      I_Contact( "状态控制数据".故障状态 )
      Coil( "状态控制数据".空闲状态 )
   END_RUNG
   RUNG wire#powerrail
      Contact( "状态控制数据".空闲状态 )
   END_RUNG wire#w1
   RUNG wire#powerrail
      Contact( "状态控制数据".空闲状态 )
      { S7_Templates := "SrcType := Int" } EQ_Contact(in1 := "三站MES读取数据".订单数据.开始信号, in2 := 1)
      Coil( "状态控制数据".忙碌状态 )
   END_RUNG
   RUNG wire#powerrail
      Contact( "初始化数据".初始化故障 )
      wire#w2
      Coil( "状态控制数据".故障状态 )
   END_RUNG
   RUNG wire#powerrail
      Contact( "初始化数据".报警总输出 )
   END_RUNG wire#w2
   // the same network as SCL:
   "状态控制数据".在线状态 := TRUE;
   IF "状态控制数据".在线状态 THEN "三站MES读取数据".三站数据.在线状态 := 1; END_IF;
   "状态控制数据".空闲状态 := ("初始化数据".初始化完成 OR "状态控制数据".空闲状态) AND NOT "初始化数据".报警总输出 AND NOT "初始化数据".急停状态 AND NOT "状态控制数据".故障状态;
   "状态控制数据".忙碌状态 := "状态控制数据".空闲状态 AND ("三站MES读取数据".订单数据.开始信号 = 1);
   "状态控制数据".故障状态 := "初始化数据".初始化故障 OR "初始化数据".报警总输出;
END_REGION

REGION Network 2: 安全光栅和急停
   RUNG wire#powerrail
      Contact( "[156]安全光栅" )
      Coil( "三站数据".安全光栅 )
   END_RUNG
   RUNG wire#powerrail
      I_Contact( "[112]急停" )
      Coil( "初始化数据".急停状态 )
   END_RUNG
   // the same network as SCL:
   "三站数据".安全光栅 := "[156]安全光栅";
   "初始化数据".急停状态 := NOT "[112]急停";
END_REGION

REGION Network 3: 三色灯————黄灯
   RUNG wire#powerrail
      Contact( "初始化数据".初始化中 )
      Contact( "Clock_0.5Hz" )
      wire#w1
      Coil( "初始化数据".黄灯_内部 )
   END_RUNG
   RUNG wire#powerrail
      Contact( "初始化数据".初始化完成 )
      I_Contact( "初始化数据".自动运行模式 )
   END_RUNG wire#w1
   // the same network as SCL:
   "初始化数据".黄灯_内部 := ("初始化数据".初始化中 AND "Clock_0.5Hz") OR ("初始化数据".初始化完成 AND NOT "初始化数据".自动运行模式);
END_REGION

REGION Network 4: 三色灯————绿灯
   RUNG wire#powerrail
      Contact( "初始化数据".自动运行模式 )
      { S7_Templates := "SrcType := Int" } EQ_Contact(in1 := "初始化数据".报警等级, in2 := 0)
      I_Contact( "状态控制数据".忙碌状态 )
      wire#w1
      Coil( "初始化数据".绿灯_内部 )
   END_RUNG
   RUNG wire#powerrail
      Contact( "初始化数据".自动运行模式 )
      { S7_Templates := "SrcType := Int" } EQ_Contact(in1 := "初始化数据".报警等级, in2 := 0)
      Contact( "状态控制数据".忙碌状态 )
      Contact( "Clock_0.5Hz" )
   END_RUNG wire#w1
   // the same network as SCL:
   "初始化数据".绿灯_内部 := ("初始化数据".自动运行模式 AND ("初始化数据".报警等级 = 0) AND NOT "状态控制数据".忙碌状态) OR ("初始化数据".自动运行模式 AND ("初始化数据".报警等级 = 0) AND "状态控制数据".忙碌状态 AND "Clock_0.5Hz");
END_REGION

REGION Network 5: 三色灯————红灯
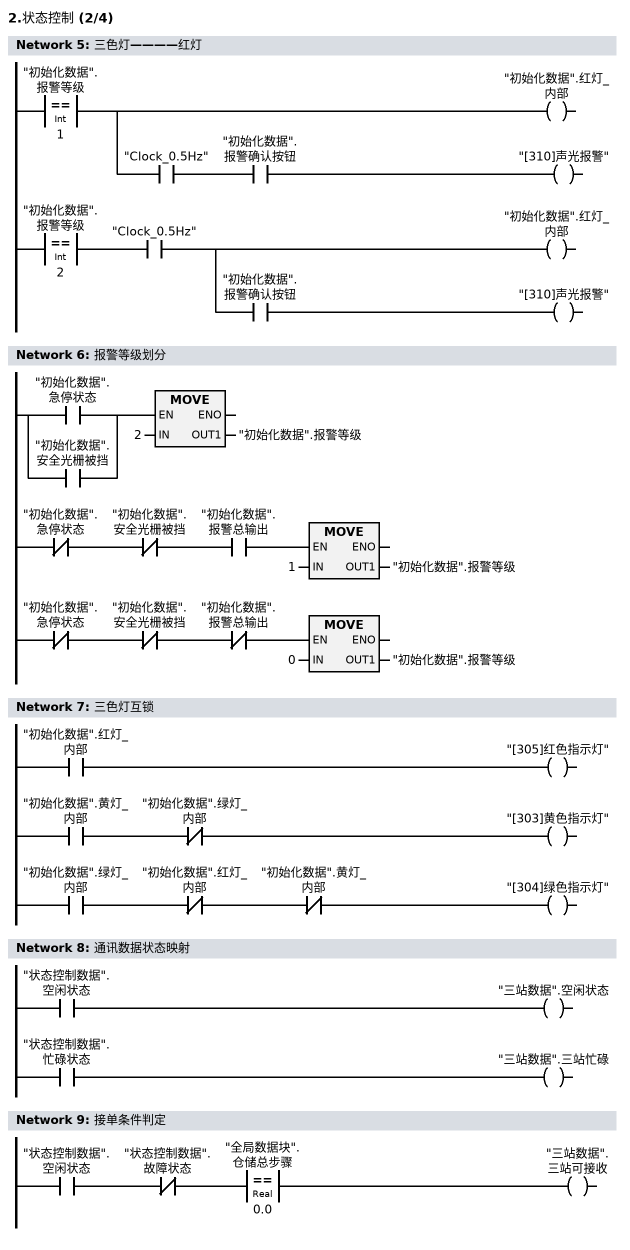
   RUNG wire#powerrail
      { S7_Templates := "SrcType := Int" } EQ_Contact(in1 := "初始化数据".报警等级, in2 := 1)
      wire#w1
      Coil( "初始化数据".红灯_内部 )
   END_RUNG
   RUNG wire#w1
      Contact( "Clock_0.5Hz" )
      Contact( "初始化数据".报警确认按钮 )
      Coil( "[310]声光报警" )
   END_RUNG
   RUNG wire#powerrail
      { S7_Templates := "SrcType := Int" } EQ_Contact(in1 := "初始化数据".报警等级, in2 := 2)
      Contact( "Clock_0.5Hz" )
      wire#w2
      Coil( "初始化数据".红灯_内部 )
   END_RUNG
   RUNG wire#w2
      Contact( "初始化数据".报警确认按钮 )
      Coil( "[310]声光报警" )
   END_RUNG
   // the same network as SCL:
   "初始化数据".红灯_内部 := "初始化数据".报警等级 = 1;
   "[310]声光报警" := "初始化数据".红灯_内部 AND "Clock_0.5Hz" AND "初始化数据".报警确认按钮;
   "初始化数据".红灯_内部 := ("初始化数据".报警等级 = 2) AND "Clock_0.5Hz";
   "[310]声光报警" := "初始化数据".红灯_内部 AND "初始化数据".报警确认按钮;
END_REGION

REGION Network 6: 报警等级划分
   RUNG wire#powerrail
      Contact( "初始化数据".急停状态 )
      wire#w1
      Move(in := 2, out1 => "初始化数据".报警等级)
   END_RUNG
   RUNG wire#powerrail
      Contact( "初始化数据".安全光栅被挡 )
   END_RUNG wire#w1
   RUNG wire#powerrail
      I_Contact( "初始化数据".急停状态 )
      I_Contact( "初始化数据".安全光栅被挡 )
      Contact( "初始化数据".报警总输出 )
      Move(in := 1, out1 => "初始化数据".报警等级)
   END_RUNG
   RUNG wire#powerrail
      I_Contact( "初始化数据".急停状态 )
      I_Contact( "初始化数据".安全光栅被挡 )
      I_Contact( "初始化数据".报警总输出 )
      Move(in := 0, out1 => "初始化数据".报警等级)
   END_RUNG
   // the same network as SCL:
   IF "初始化数据".急停状态 OR "初始化数据".安全光栅被挡 THEN "初始化数据".报警等级 := 2; END_IF;
   IF NOT "初始化数据".急停状态 AND NOT "初始化数据".安全光栅被挡 AND "初始化数据".报警总输出 THEN "初始化数据".报警等级 := 1; END_IF;
   IF NOT "初始化数据".急停状态 AND NOT "初始化数据".安全光栅被挡 AND NOT "初始化数据".报警总输出 THEN "初始化数据".报警等级 := 0; END_IF;
END_REGION

REGION Network 7: 三色灯互锁
   RUNG wire#powerrail
      Contact( "初始化数据".红灯_内部 )
      Coil( "[305]红色指示灯" )
   END_RUNG
   RUNG wire#powerrail
      Contact( "初始化数据".黄灯_内部 )
      I_Contact( "初始化数据".绿灯_内部 )
      Coil( "[303]黄色指示灯" )
   END_RUNG
   RUNG wire#powerrail
      Contact( "初始化数据".绿灯_内部 )
      I_Contact( "初始化数据".红灯_内部 )
      I_Contact( "初始化数据".黄灯_内部 )
      Coil( "[304]绿色指示灯" )
   END_RUNG
   // the same network as SCL:
   "[305]红色指示灯" := "初始化数据".红灯_内部;
   "[303]黄色指示灯" := "初始化数据".黄灯_内部 AND NOT "初始化数据".绿灯_内部;
   "[304]绿色指示灯" := "初始化数据".绿灯_内部 AND NOT "初始化数据".红灯_内部 AND NOT "初始化数据".黄灯_内部;
END_REGION

REGION Network 8: 通讯数据状态映射
   RUNG wire#powerrail
      Contact( "状态控制数据".空闲状态 )
      Coil( "三站数据".空闲状态 )
   END_RUNG
   RUNG wire#powerrail
      Contact( "状态控制数据".忙碌状态 )
      Coil( "三站数据".三站忙碌 )
   END_RUNG
   // the same network as SCL:
   "三站数据".空闲状态 := "状态控制数据".空闲状态;
   "三站数据".三站忙碌 := "状态控制数据".忙碌状态;
END_REGION

REGION Network 9: 接单条件判定
   RUNG wire#powerrail
      Contact( "状态控制数据".空闲状态 )
      I_Contact( "状态控制数据".故障状态 )
      { S7_Templates := "SrcType := Real" } EQ_Contact(in1 := "全局数据块".仓储总步骤, in2 := 0.0)
      Coil( "三站数据".三站可接收 )
   END_RUNG
   // the same network as SCL:
   "三站数据".三站可接收 := "状态控制数据".空闲状态 AND NOT "状态控制数据".故障状态 AND ("全局数据块".仓储总步骤 = 0.0);
END_REGION

REGION Network 10: MES通讯数据
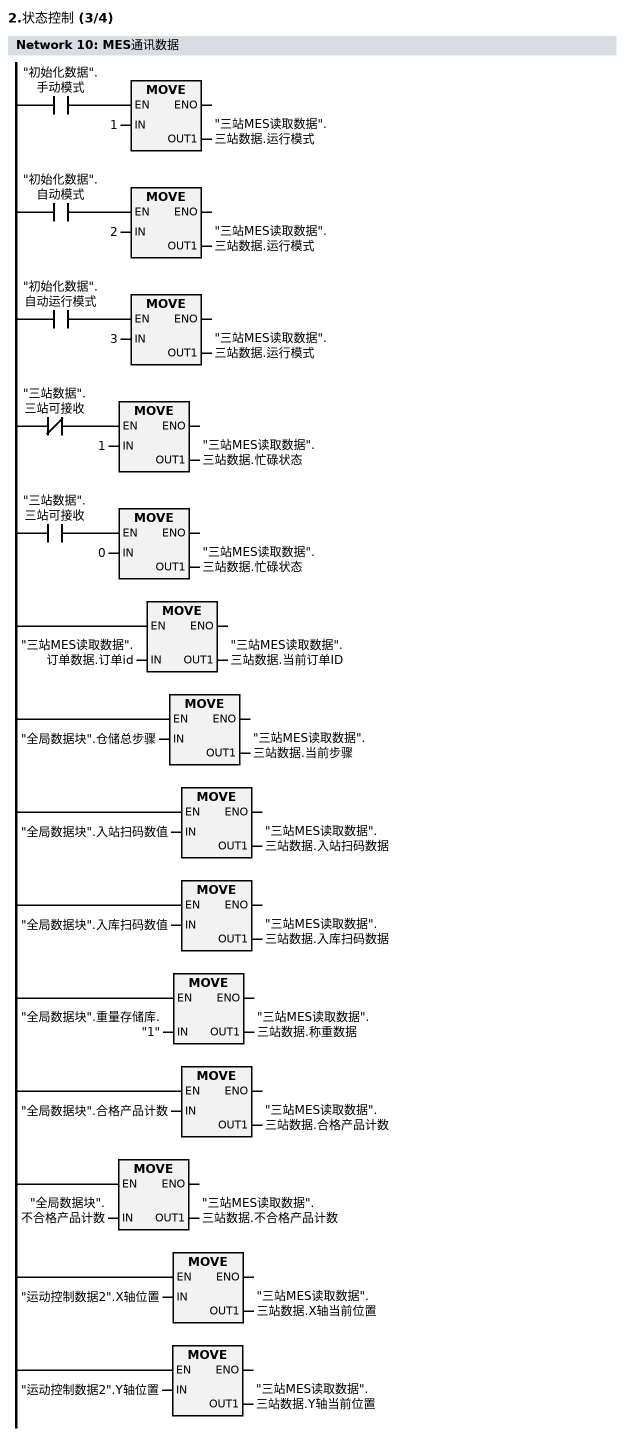
   RUNG wire#powerrail
      Contact( "初始化数据".手动模式 )
      Move(in := 1, out1 => "三站MES读取数据".三站数据.运行模式)
   END_RUNG
   RUNG wire#powerrail
      Contact( "初始化数据".自动模式 )
      Move(in := 2, out1 => "三站MES读取数据".三站数据.运行模式)
   END_RUNG
   RUNG wire#powerrail
      Contact( "初始化数据".自动运行模式 )
      Move(in := 3, out1 => "三站MES读取数据".三站数据.运行模式)
   END_RUNG
   RUNG wire#powerrail
      I_Contact( "三站数据".三站可接收 )
      Move(in := 1, out1 => "三站MES读取数据".三站数据.忙碌状态)
   END_RUNG
   RUNG wire#powerrail
      Contact( "三站数据".三站可接收 )
      Move(in := 0, out1 => "三站MES读取数据".三站数据.忙碌状态)
   END_RUNG
   RUNG wire#powerrail
      Move(in := "三站MES读取数据".订单数据.订单id, out1 => "三站MES读取数据".三站数据.当前订单ID)
   END_RUNG
   RUNG wire#powerrail
      Move(in := "全局数据块".仓储总步骤, out1 => "三站MES读取数据".三站数据.当前步骤)
   END_RUNG
   RUNG wire#powerrail
      Move(in := "全局数据块".入站扫码数值, out1 => "三站MES读取数据".三站数据.入站扫码数据)
   END_RUNG
   RUNG wire#powerrail
      Move(in := "全局数据块".入库扫码数值, out1 => "三站MES读取数据".三站数据.入库扫码数据)
   END_RUNG
   RUNG wire#powerrail
      Move(in := "全局数据块".重量存储库."1", out1 => "三站MES读取数据".三站数据.称重数据)
   END_RUNG
   RUNG wire#powerrail
      Move(in := "全局数据块".合格产品计数, out1 => "三站MES读取数据".三站数据.合格产品计数)
   END_RUNG
   RUNG wire#powerrail
      Move(in := "全局数据块".不合格产品计数, out1 => "三站MES读取数据".三站数据.不合格产品计数)
   END_RUNG
   RUNG wire#powerrail
      Move(in := "运动控制数据2".X轴位置, out1 => "三站MES读取数据".三站数据.X轴当前位置)
   END_RUNG
   RUNG wire#powerrail
      Move(in := "运动控制数据2".Y轴位置, out1 => "三站MES读取数据".三站数据.Y轴当前位置)
   END_RUNG
   // the same network as SCL:
   IF "初始化数据".手动模式 THEN "三站MES读取数据".三站数据.运行模式 := 1; END_IF;
   IF "初始化数据".自动模式 THEN "三站MES读取数据".三站数据.运行模式 := 2; END_IF;
   IF "初始化数据".自动运行模式 THEN "三站MES读取数据".三站数据.运行模式 := 3; END_IF;
   IF NOT "三站数据".三站可接收 THEN "三站MES读取数据".三站数据.忙碌状态 := 1; END_IF;
   IF "三站数据".三站可接收 THEN "三站MES读取数据".三站数据.忙碌状态 := 0; END_IF;
   "三站MES读取数据".三站数据.当前订单ID := "三站MES读取数据".订单数据.订单id;
   "三站MES读取数据".三站数据.当前步骤 := "全局数据块".仓储总步骤;
   "三站MES读取数据".三站数据.入站扫码数据 := "全局数据块".入站扫码数值;
   "三站MES读取数据".三站数据.入库扫码数据 := "全局数据块".入库扫码数值;
   "三站MES读取数据".三站数据.称重数据 := "全局数据块".重量存储库."1";
   "三站MES读取数据".三站数据.合格产品计数 := "全局数据块".合格产品计数;
   "三站MES读取数据".三站数据.不合格产品计数 := "全局数据块".不合格产品计数;
   "三站MES读取数据".三站数据.X轴当前位置 := "运动控制数据2".X轴位置;
   "三站MES读取数据".三站数据.Y轴当前位置 := "运动控制数据2".Y轴位置;
END_REGION

REGION Network 11
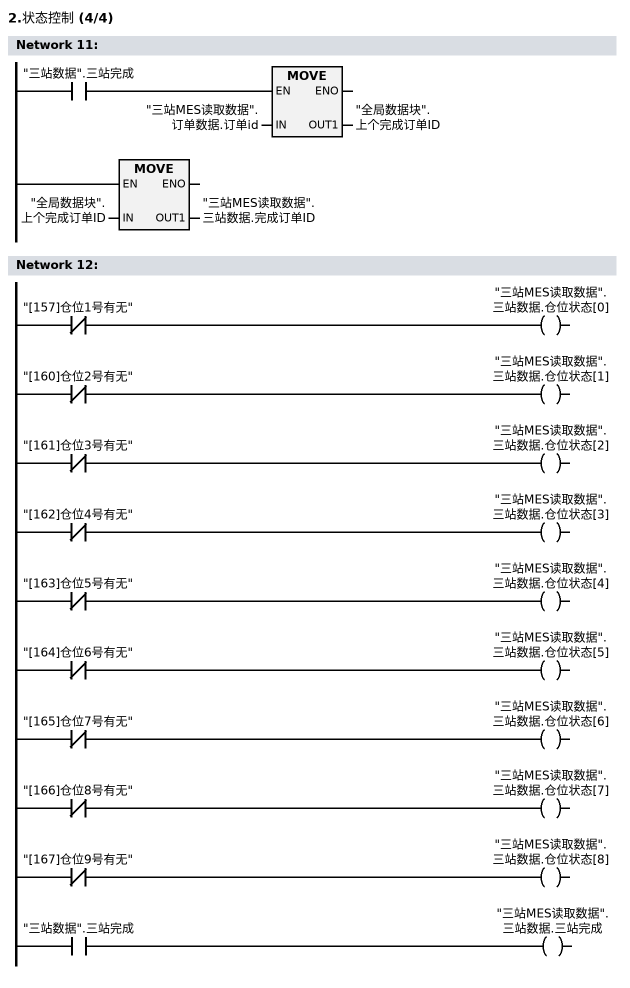
   RUNG wire#powerrail
      Contact( "三站数据".三站完成 )
      Move(in := "三站MES读取数据".订单数据.订单id, out1 => "全局数据块".上个完成订单ID)
   END_RUNG
   RUNG wire#powerrail
      Move(in := "全局数据块".上个完成订单ID, out1 => "三站MES读取数据".三站数据.完成订单ID)
   END_RUNG
   // the same network as SCL:
   IF "三站数据".三站完成 THEN "全局数据块".上个完成订单ID := "三站MES读取数据".订单数据.订单id; END_IF;
   "三站MES读取数据".三站数据.完成订单ID := "全局数据块".上个完成订单ID;
END_REGION

REGION Network 12
   RUNG wire#powerrail
      I_Contact( "[157]仓位1号有无" )
      Coil( "三站MES读取数据".三站数据.仓位状态[0] )
   END_RUNG
   RUNG wire#powerrail
      I_Contact( "[160]仓位2号有无" )
      Coil( "三站MES读取数据".三站数据.仓位状态[1] )
   END_RUNG
   RUNG wire#powerrail
      I_Contact( "[161]仓位3号有无" )
      Coil( "三站MES读取数据".三站数据.仓位状态[2] )
   END_RUNG
   RUNG wire#powerrail
      I_Contact( "[162]仓位4号有无" )
      Coil( "三站MES读取数据".三站数据.仓位状态[3] )
   END_RUNG
   RUNG wire#powerrail
      I_Contact( "[163]仓位5号有无" )
      Coil( "三站MES读取数据".三站数据.仓位状态[4] )
   END_RUNG
   RUNG wire#powerrail
      I_Contact( "[164]仓位6号有无" )
      Coil( "三站MES读取数据".三站数据.仓位状态[5] )
   END_RUNG
   RUNG wire#powerrail
      I_Contact( "[165]仓位7号有无" )
      Coil( "三站MES读取数据".三站数据.仓位状态[6] )
   END_RUNG
   RUNG wire#powerrail
      I_Contact( "[166]仓位8号有无" )
      Coil( "三站MES读取数据".三站数据.仓位状态[7] )
   END_RUNG
   RUNG wire#powerrail
      I_Contact( "[167]仓位9号有无" )
      Coil( "三站MES读取数据".三站数据.仓位状态[8] )
   END_RUNG
   RUNG wire#powerrail
      Contact( "三站数据".三站完成 )
      Coil( "三站MES读取数据".三站数据.三站完成 )
   END_RUNG
   // the same network as SCL:
   "三站MES读取数据".三站数据.仓位状态[0] := NOT "[157]仓位1号有无";
   "三站MES读取数据".三站数据.仓位状态[1] := NOT "[160]仓位2号有无";
   "三站MES读取数据".三站数据.仓位状态[2] := NOT "[161]仓位3号有无";
   "三站MES读取数据".三站数据.仓位状态[3] := NOT "[162]仓位4号有无";
   "三站MES读取数据".三站数据.仓位状态[4] := NOT "[163]仓位5号有无";
   "三站MES读取数据".三站数据.仓位状态[5] := NOT "[164]仓位6号有无";
   "三站MES读取数据".三站数据.仓位状态[6] := NOT "[165]仓位7号有无";
   "三站MES读取数据".三站数据.仓位状态[7] := NOT "[166]仓位8号有无";
   "三站MES读取数据".三站数据.仓位状态[8] := NOT "[167]仓位9号有无";
   "三站MES读取数据".三站数据.三站完成 := "三站数据".三站完成;
END_REGION
END_FUNCTION

FUNCTION "1.报警程序" : Void   // FC14, LAD
{ S7_Optimized_Access := 'TRUE' }
VERSION : 0.1
BEGIN
END_FUNCTION

FUNCTION "测试" : Void   // FC16, LAD
{ S7_Optimized_Access := 'TRUE' }
VERSION : 0.1
BEGIN
END_FUNCTION

FUNCTION "手动模式流程" : Void   // FC19, LAD
{ S7_Optimized_Access := 'TRUE' }
VERSION : 0.1
   VAR_TEMP   // added for the SCL form of the ladder/FBD networks
      _w1 : Bool;
      _w2 : Bool;
      _w3 : Bool;
      _w4 : Bool;
   END_VAR
BEGIN

REGION Network 1
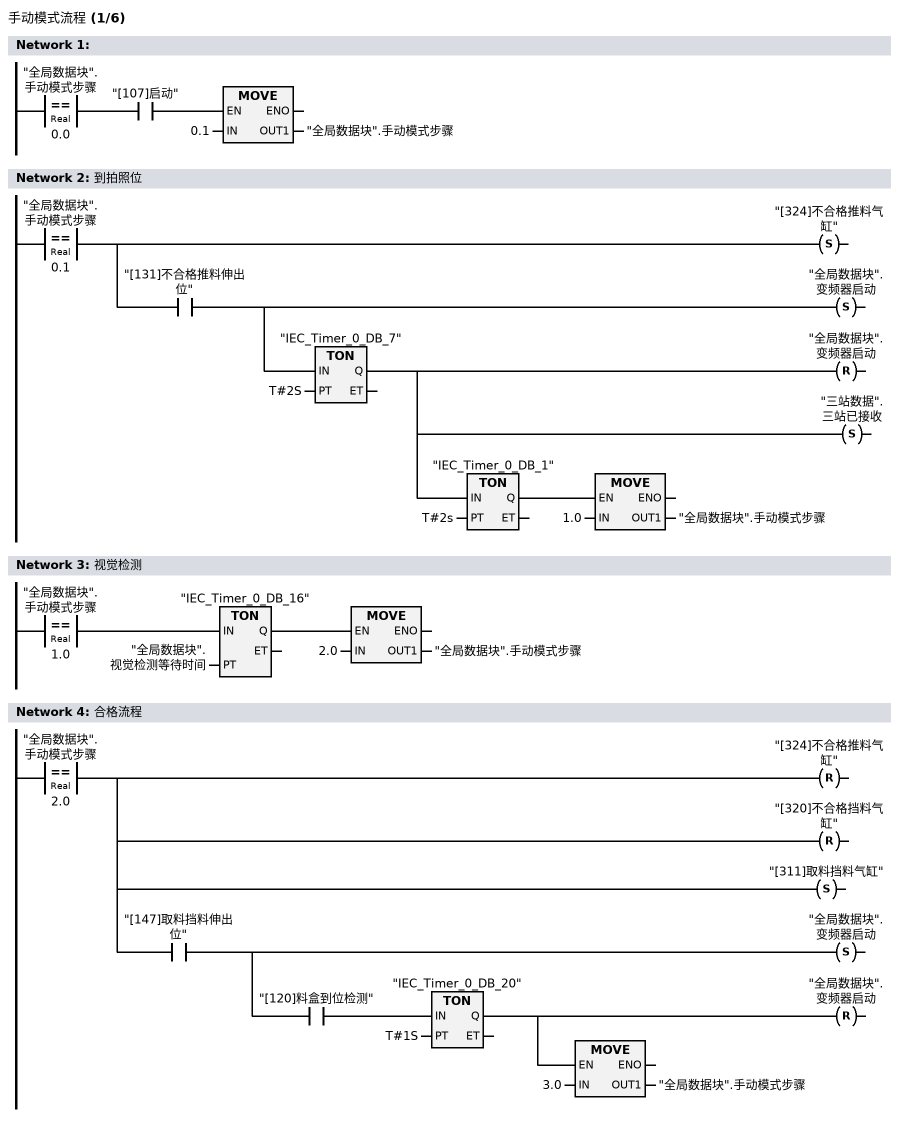
   RUNG wire#powerrail
      { S7_Templates := "SrcType := Real" } EQ_Contact(in1 := "全局数据块".手动模式步骤, in2 := 0.0)
      Contact( "[107]启动" )
      Move(in := 0.1, out1 => "全局数据块".手动模式步骤)
   END_RUNG
   // the same network as SCL:
   IF ("全局数据块".手动模式步骤 = 0.0) AND "[107]启动" THEN "全局数据块".手动模式步骤 := 0.1; END_IF;
END_REGION

REGION Network 2: 到拍照位
   #_w1 := "全局数据块".手动模式步骤 = 0.1;
   IF #_w1 THEN "[324]不合格推料气缸" := TRUE; END_IF;
   #_w2 := #_w1 AND "[131]不合格推料伸出位";
   IF #_w2 THEN "全局数据块".变频器启动 := TRUE; END_IF;
   "IEC_Timer_0_DB_7".TON(IN := #_w2, PT := T#2S);
   IF "IEC_Timer_0_DB_7".Q THEN
       "全局数据块".变频器启动 := FALSE;
       "三站数据".三站已接收 := TRUE;
   END_IF;
   "IEC_Timer_0_DB_1".TON(IN := "IEC_Timer_0_DB_7".Q, PT := T#2s);
   IF "IEC_Timer_0_DB_1".Q THEN "全局数据块".手动模式步骤 := 1.0; END_IF;
END_REGION

REGION Network 3: 视觉检测
   "IEC_Timer_0_DB_16".TON(IN := "全局数据块".手动模式步骤 = 1.0, PT := "全局数据块".视觉检测等待时间);
   IF "IEC_Timer_0_DB_16".Q THEN "全局数据块".手动模式步骤 := 2.0; END_IF;
END_REGION

REGION Network 4: 合格流程
   #_w1 := "全局数据块".手动模式步骤 = 2.0;
   IF #_w1 THEN
       "[324]不合格推料气缸" := FALSE;
       "[320]不合格挡料气缸" := FALSE;
       "[311]取料挡料气缸" := TRUE;
   END_IF;
   #_w2 := #_w1 AND "[147]取料挡料伸出位";
   IF #_w2 THEN "全局数据块".变频器启动 := TRUE; END_IF;
   "IEC_Timer_0_DB_20".TON(IN := #_w2 AND "[120]料盒到位检测", PT := T#1S);
   IF "IEC_Timer_0_DB_20".Q THEN
       "全局数据块".变频器启动 := FALSE;
       "全局数据块".手动模式步骤 := 3.0;
   END_IF;
END_REGION

REGION Network 5: 不合格流程
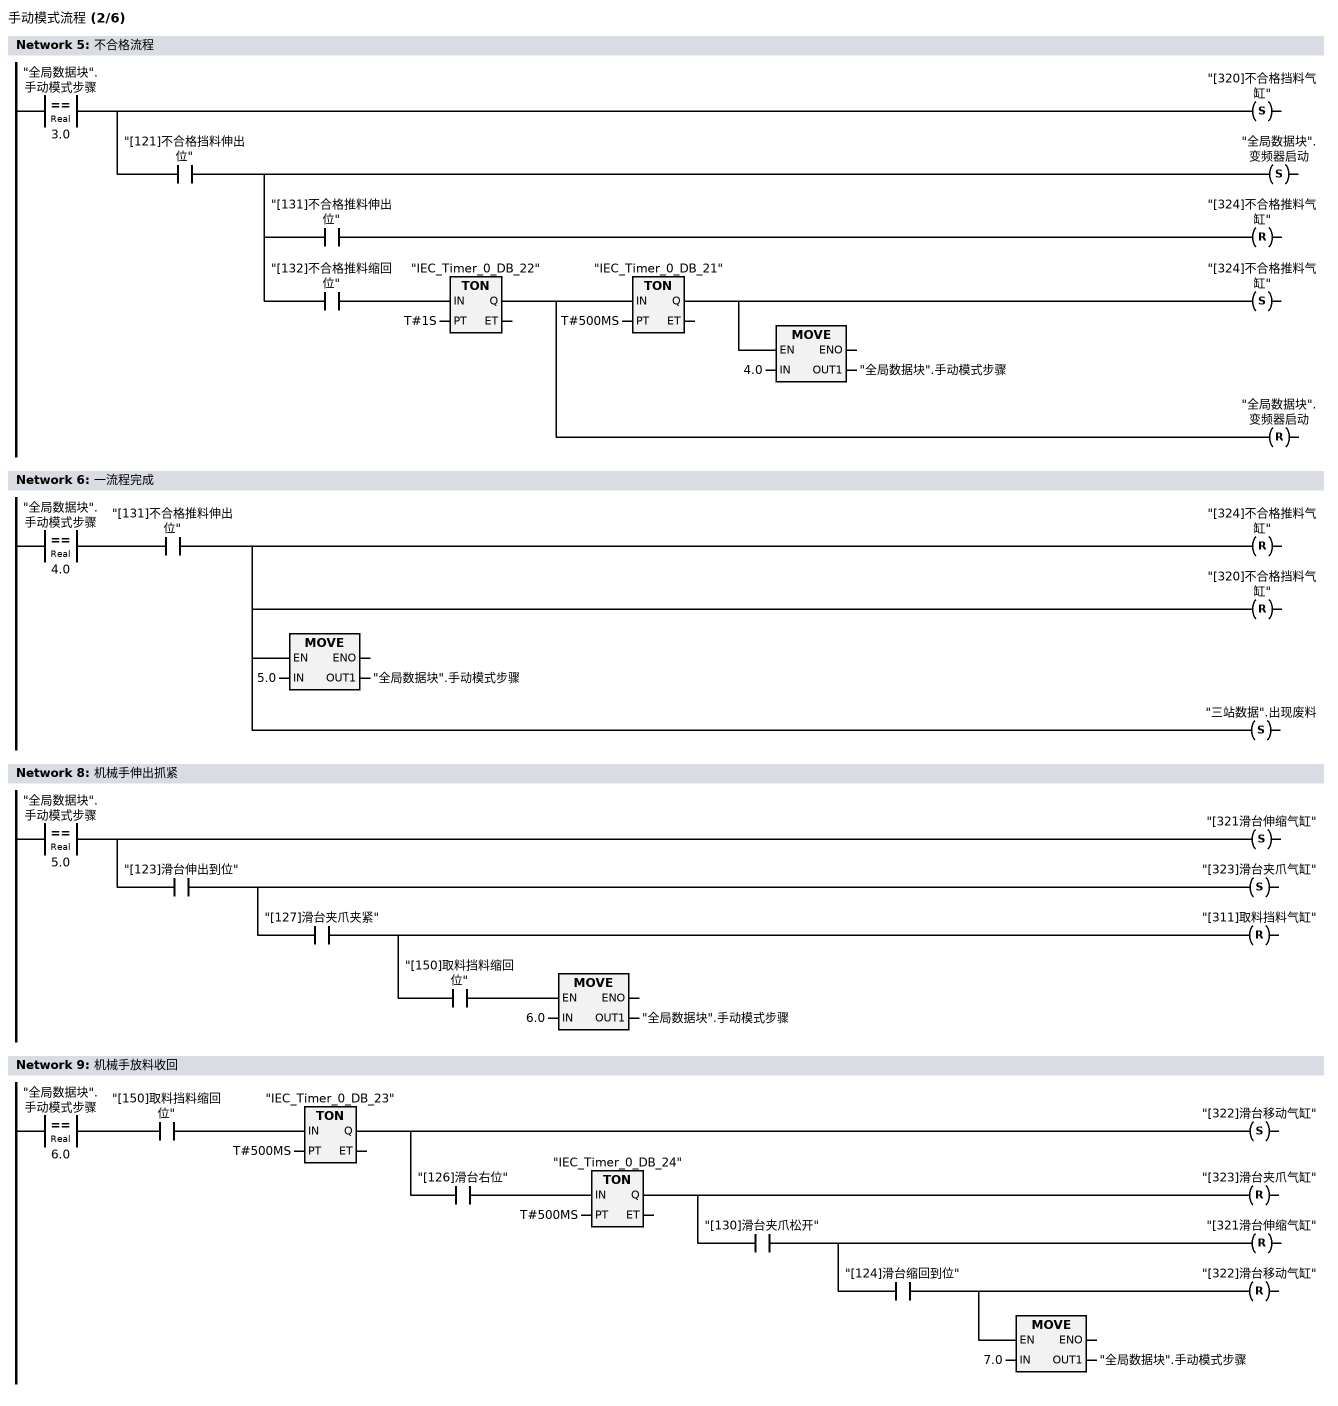
   #_w1 := "全局数据块".手动模式步骤 = 3.0;
   IF #_w1 THEN "[320]不合格挡料气缸" := TRUE; END_IF;
   #_w2 := #_w1 AND "[121]不合格挡料伸出位";
   IF #_w2 THEN "全局数据块".变频器启动 := TRUE; END_IF;
   IF #_w2 AND "[131]不合格推料伸出位" THEN "[324]不合格推料气缸" := FALSE; END_IF;
   "IEC_Timer_0_DB_22".TON(IN := #_w2 AND "[132]不合格推料缩回位", PT := T#1S);
   "IEC_Timer_0_DB_21".TON(IN := "IEC_Timer_0_DB_22".Q, PT := T#500MS);
   IF "IEC_Timer_0_DB_21".Q THEN
       "[324]不合格推料气缸" := TRUE;
       "全局数据块".手动模式步骤 := 4.0;
   END_IF;
   IF "IEC_Timer_0_DB_22".Q THEN "全局数据块".变频器启动 := FALSE; END_IF;
END_REGION

REGION Network 6: 一流程完成
   RUNG wire#powerrail
      { S7_Templates := "SrcType := Real" } EQ_Contact(in1 := "全局数据块".手动模式步骤, in2 := 4.0)
      Contact( "[131]不合格推料伸出位" )
      wire#w1
      R_Coil( "[324]不合格推料气缸" )
   END_RUNG
   RUNG wire#w1
      R_Coil( "[320]不合格挡料气缸" )
   END_RUNG
   RUNG wire#w1
      Move(in := 5.0, out1 => "全局数据块".手动模式步骤)
   END_RUNG
   RUNG wire#w1
      S_Coil( "三站数据".出现废料 )
   END_RUNG
   // the same network as SCL:
   #_w1 := ("全局数据块".手动模式步骤 = 4.0) AND "[131]不合格推料伸出位";
   IF #_w1 THEN
       "[324]不合格推料气缸" := FALSE;
       "[320]不合格挡料气缸" := FALSE;
       "全局数据块".手动模式步骤 := 5.0;
       "三站数据".出现废料 := TRUE;
   END_IF;
END_REGION

REGION Network 7: 开始二流程
END_REGION

REGION Network 8: 机械手伸出抓紧
   RUNG wire#powerrail
      { S7_Templates := "SrcType := Real" } EQ_Contact(in1 := "全局数据块".手动模式步骤, in2 := 5.0)
      wire#w1
      S_Coil( "[321滑台伸缩气缸" )
   END_RUNG
   RUNG wire#w1
      Contact( "[123]滑台伸出到位" )
      wire#w2
      S_Coil( "[323]滑台夹爪气缸" )
   END_RUNG
   RUNG wire#w2
      Contact( "[127]滑台夹爪夹紧" )
      wire#w3
      R_Coil( "[311]取料挡料气缸" )
   END_RUNG
   RUNG wire#w3
      Contact( "[150]取料挡料缩回位" )
      Move(in := 6.0, out1 => "全局数据块".手动模式步骤)
   END_RUNG
   // the same network as SCL:
   #_w1 := "全局数据块".手动模式步骤 = 5.0;
   IF #_w1 THEN "[321滑台伸缩气缸" := TRUE; END_IF;
   #_w2 := #_w1 AND "[123]滑台伸出到位";
   IF #_w2 THEN "[323]滑台夹爪气缸" := TRUE; END_IF;
   #_w3 := #_w2 AND "[127]滑台夹爪夹紧";
   IF #_w3 THEN "[311]取料挡料气缸" := FALSE; END_IF;
   IF #_w3 AND "[150]取料挡料缩回位" THEN "全局数据块".手动模式步骤 := 6.0; END_IF;
END_REGION

REGION Network 9: 机械手放料收回
   "IEC_Timer_0_DB_23".TON(IN := ("全局数据块".手动模式步骤 = 6.0) AND "[150]取料挡料缩回位", PT := T#500MS);
   IF "IEC_Timer_0_DB_23".Q THEN "[322]滑台移动气缸" := TRUE; END_IF;
   "IEC_Timer_0_DB_24".TON(IN := "IEC_Timer_0_DB_23".Q AND "[126]滑台右位", PT := T#500MS);
   IF "IEC_Timer_0_DB_24".Q THEN "[323]滑台夹爪气缸" := FALSE; END_IF;
   #_w1 := "IEC_Timer_0_DB_24".Q AND "[130]滑台夹爪松开";
   IF #_w1 THEN "[321滑台伸缩气缸" := FALSE; END_IF;
   #_w2 := #_w1 AND "[124]滑台缩回到位";
   IF #_w2 THEN
       "[322]滑台移动气缸" := FALSE;
       "全局数据块".手动模式步骤 := 7.0;
   END_IF;
END_REGION

REGION Network 10: 称重
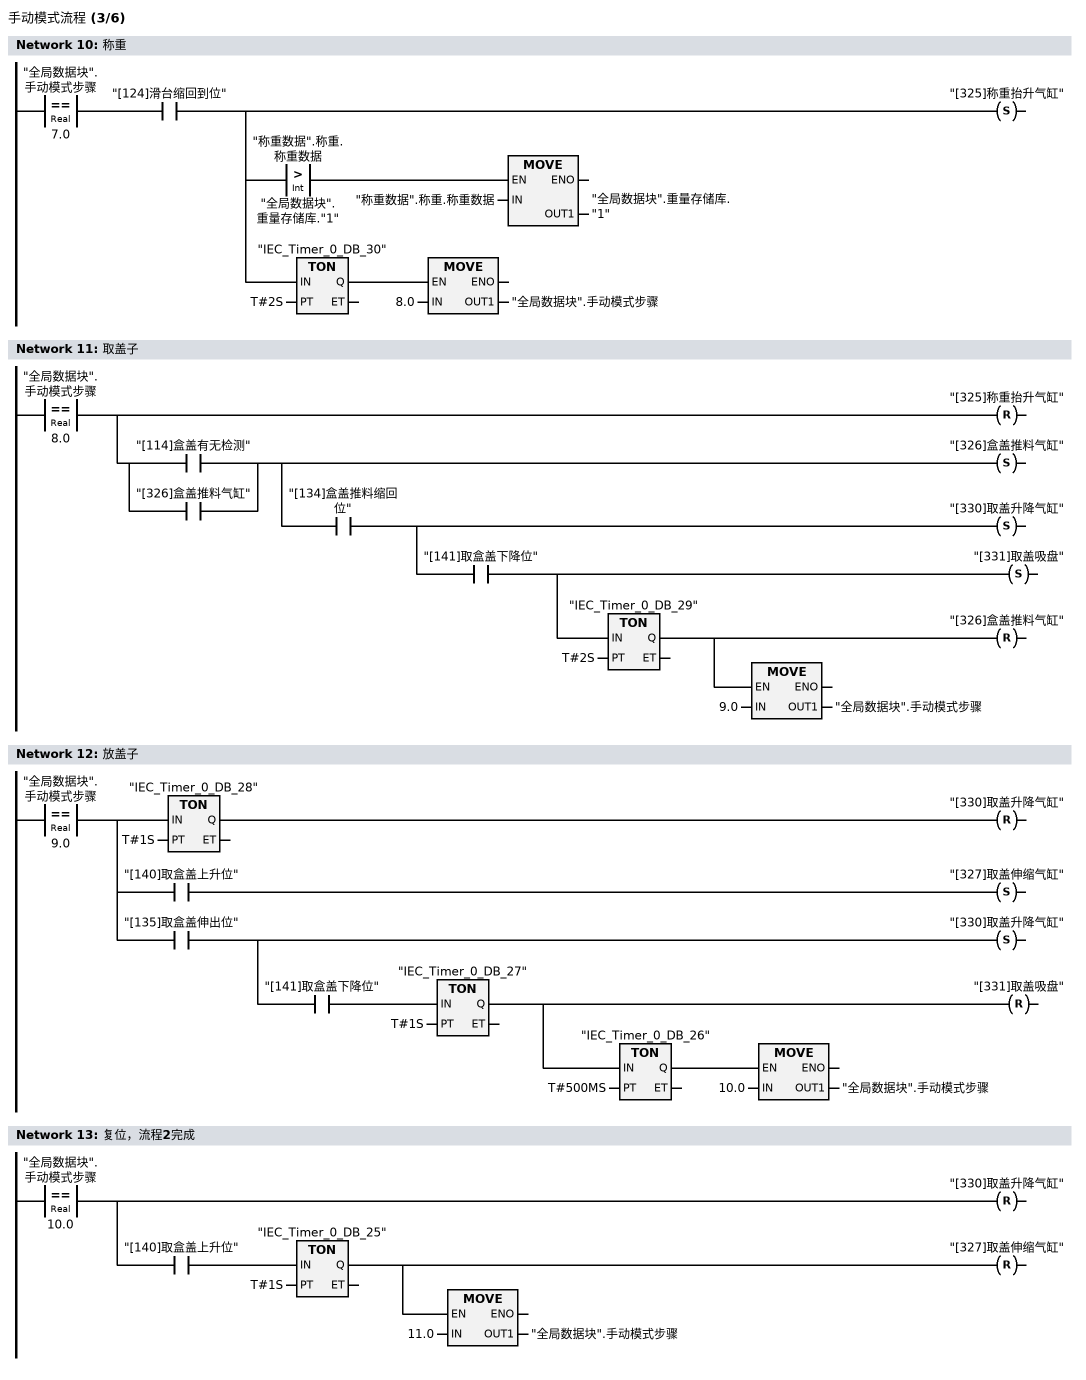
   #_w1 := ("全局数据块".手动模式步骤 = 7.0) AND "[124]滑台缩回到位";
   IF #_w1 THEN "[325]称重抬升气缸" := TRUE; END_IF;
   IF #_w1 AND ("称重数据".称重.称重数据 > "全局数据块".重量存储库."1") THEN "全局数据块".重量存储库."1" := "称重数据".称重.称重数据; END_IF;
   "IEC_Timer_0_DB_30".TON(IN := #_w1, PT := T#2S);
   IF "IEC_Timer_0_DB_30".Q THEN "全局数据块".手动模式步骤 := 8.0; END_IF;
END_REGION

REGION Network 11: 取盖子
   #_w1 := "全局数据块".手动模式步骤 = 8.0;
   IF #_w1 THEN "[325]称重抬升气缸" := FALSE; END_IF;
   #_w2 := #_w1 AND ("[114]盒盖有无检测" OR "[326]盒盖推料气缸");
   IF #_w2 THEN "[326]盒盖推料气缸" := TRUE; END_IF;
   #_w3 := #_w2 AND "[134]盒盖推料缩回位";
   IF #_w3 THEN "[330]取盖升降气缸" := TRUE; END_IF;
   #_w4 := #_w3 AND "[141]取盒盖下降位";
   IF #_w4 THEN "[331]取盖吸盘" := TRUE; END_IF;
   "IEC_Timer_0_DB_29".TON(IN := #_w4, PT := T#2S);
   IF "IEC_Timer_0_DB_29".Q THEN
       "[326]盒盖推料气缸" := FALSE;
       "全局数据块".手动模式步骤 := 9.0;
   END_IF;
END_REGION

REGION Network 12: 放盖子
   #_w1 := "全局数据块".手动模式步骤 = 9.0;
   "IEC_Timer_0_DB_28".TON(IN := #_w1, PT := T#1S);
   IF "IEC_Timer_0_DB_28".Q THEN "[330]取盖升降气缸" := FALSE; END_IF;
   IF #_w1 AND "[140]取盒盖上升位" THEN "[327]取盖伸缩气缸" := TRUE; END_IF;
   #_w2 := #_w1 AND "[135]取盒盖伸出位";
   IF #_w2 THEN "[330]取盖升降气缸" := TRUE; END_IF;
   "IEC_Timer_0_DB_27".TON(IN := #_w2 AND "[141]取盒盖下降位", PT := T#1S);
   IF "IEC_Timer_0_DB_27".Q THEN "[331]取盖吸盘" := FALSE; END_IF;
   "IEC_Timer_0_DB_26".TON(IN := "IEC_Timer_0_DB_27".Q, PT := T#500MS);
   IF "IEC_Timer_0_DB_26".Q THEN "全局数据块".手动模式步骤 := 10.0; END_IF;
END_REGION

REGION Network 13: 复位，流程2完成
   #_w1 := "全局数据块".手动模式步骤 = 10.0;
   IF #_w1 THEN "[330]取盖升降气缸" := FALSE; END_IF;
   "IEC_Timer_0_DB_25".TON(IN := #_w1 AND "[140]取盒盖上升位", PT := T#1S);
   IF "IEC_Timer_0_DB_25".Q THEN
       "[327]取盖伸缩气缸" := FALSE;
       "全局数据块".手动模式步骤 := 11.0;
   END_IF;
END_REGION

REGION Network 14: 到取料位
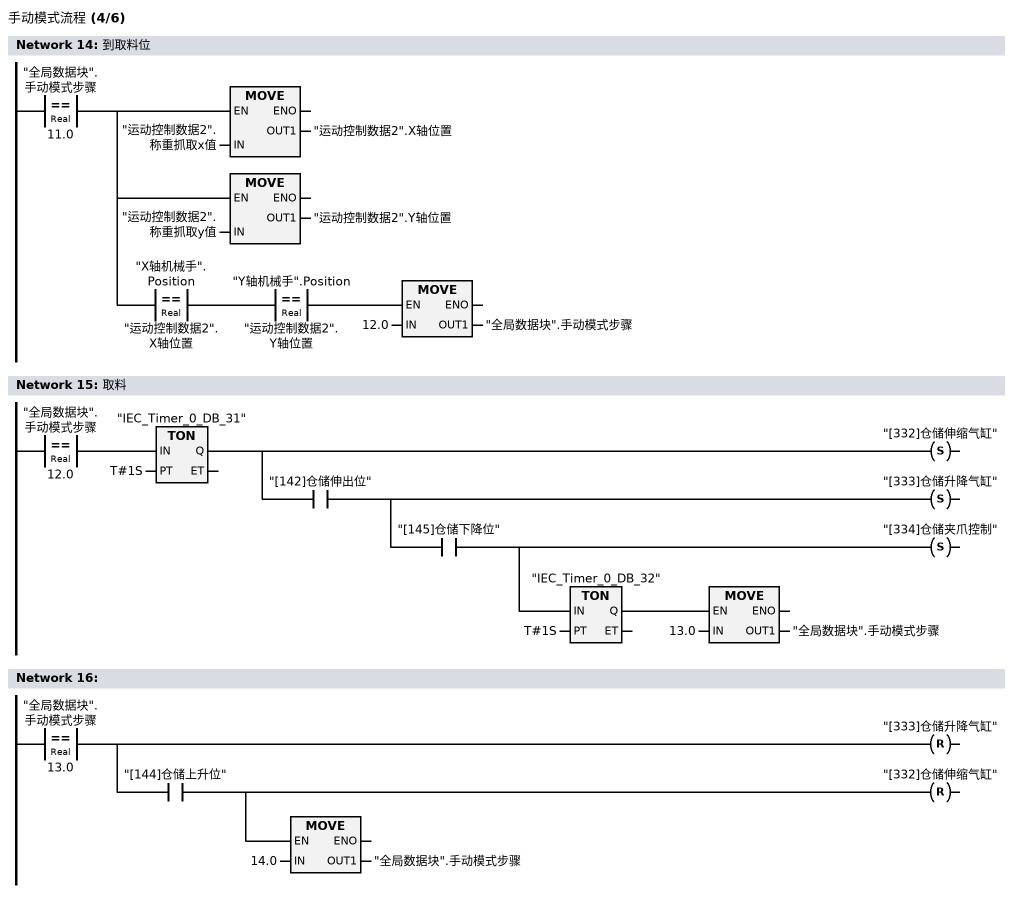
   RUNG wire#powerrail
      { S7_Templates := "SrcType := Real" } EQ_Contact(in1 := "全局数据块".手动模式步骤, in2 := 11.0)
      wire#w1
      Move(in := "运动控制数据2".称重抓取x值, out1 => "运动控制数据2".X轴位置)
   END_RUNG
   RUNG wire#w1
      Move(in := "运动控制数据2".称重抓取y值, out1 => "运动控制数据2".Y轴位置)
   END_RUNG
   RUNG wire#w1
      { S7_Templates := "SrcType := Real" } EQ_Contact(in1 := "X轴机械手".Position, in2 := "运动控制数据2".X轴位置)
      { S7_Templates := "SrcType := Real" } EQ_Contact(in1 := "Y轴机械手".Position, in2 := "运动控制数据2".Y轴位置)
      Move(in := 12.0, out1 => "全局数据块".手动模式步骤)
   END_RUNG
   // the same network as SCL:
   #_w1 := "全局数据块".手动模式步骤 = 11.0;
   IF #_w1 THEN
       "运动控制数据2".X轴位置 := "运动控制数据2".称重抓取x值;
       "运动控制数据2".Y轴位置 := "运动控制数据2".称重抓取y值;
   END_IF;
   IF #_w1 AND ("X轴机械手".Position = "运动控制数据2".X轴位置) AND ("Y轴机械手".Position = "运动控制数据2".Y轴位置) THEN
       "全局数据块".手动模式步骤 := 12.0;
   END_IF;
END_REGION

REGION Network 15: 取料
   "IEC_Timer_0_DB_31".TON(IN := "全局数据块".手动模式步骤 = 12.0, PT := T#1S);
   IF "IEC_Timer_0_DB_31".Q THEN "[332]仓储伸缩气缸" := TRUE; END_IF;
   #_w1 := "IEC_Timer_0_DB_31".Q AND "[142]仓储伸出位";
   IF #_w1 THEN "[333]仓储升降气缸" := TRUE; END_IF;
   #_w2 := #_w1 AND "[145]仓储下降位";
   IF #_w2 THEN "[334]仓储夹爪控制" := TRUE; END_IF;
   "IEC_Timer_0_DB_32".TON(IN := #_w2, PT := T#1S);
   IF "IEC_Timer_0_DB_32".Q THEN "全局数据块".手动模式步骤 := 13.0; END_IF;
END_REGION

REGION Network 16
   RUNG wire#powerrail
      { S7_Templates := "SrcType := Real" } EQ_Contact(in1 := "全局数据块".手动模式步骤, in2 := 13.0)
      wire#w1
      R_Coil( "[333]仓储升降气缸" )
   END_RUNG
   RUNG wire#w1
      Contact( "[144]仓储上升位" )
      wire#w2
      R_Coil( "[332]仓储伸缩气缸" )
   END_RUNG
   RUNG wire#w2
      Move(in := 14.0, out1 => "全局数据块".手动模式步骤)
   END_RUNG
   // the same network as SCL:
   #_w1 := "全局数据块".手动模式步骤 = 13.0;
   IF #_w1 THEN "[333]仓储升降气缸" := FALSE; END_IF;
   #_w2 := #_w1 AND "[144]仓储上升位";
   IF #_w2 THEN
       "[332]仓储伸缩气缸" := FALSE;
       "全局数据块".手动模式步骤 := 14.0;
   END_IF;
END_REGION

REGION Network 17: 仓位选择
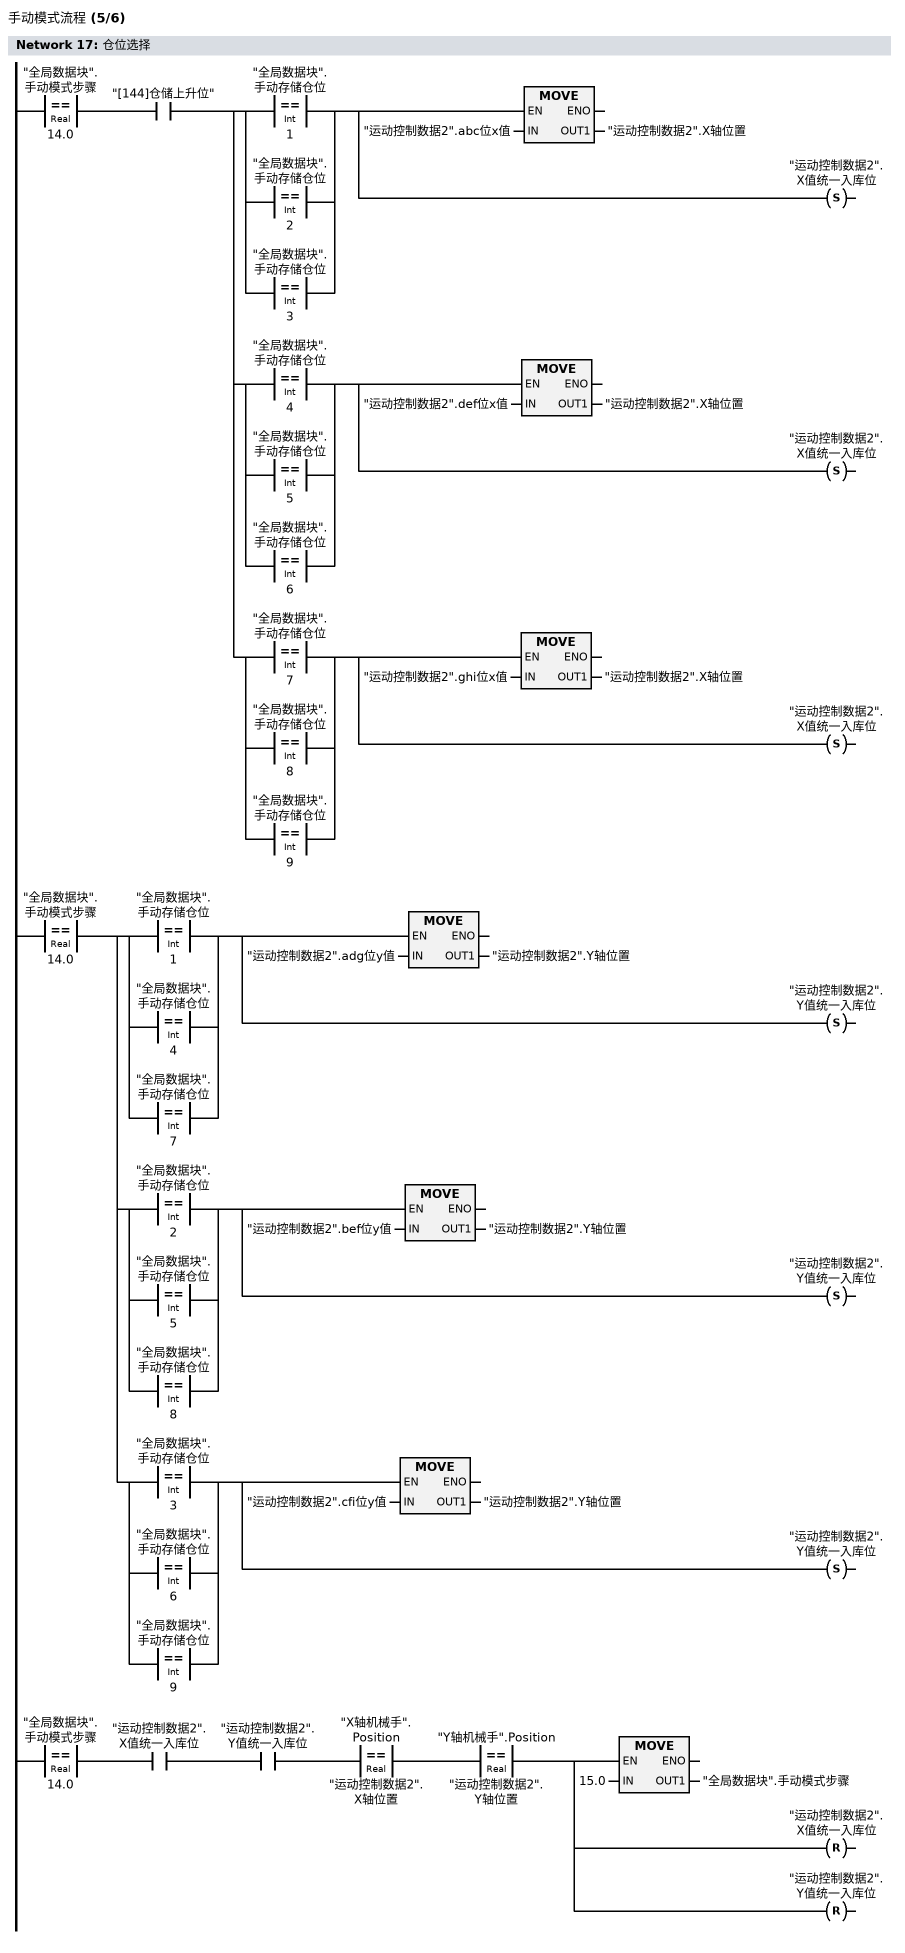
   RUNG wire#powerrail
      { S7_Templates := "SrcType := Real" } EQ_Contact(in1 := "全局数据块".手动模式步骤, in2 := 14.0)
      Contact( "[144]仓储上升位" )
      wire#w1
      { S7_Templates := "SrcType := Int" } EQ_Contact(in1 := "全局数据块".手动存储仓位, in2 := 1)
      wire#w2
      Move(in := "运动控制数据2".abc位x值, out1 => "运动控制数据2".X轴位置)
   END_RUNG
   RUNG wire#w1
      { S7_Templates := "SrcType := Int" } EQ_Contact(in1 := "全局数据块".手动存储仓位, in2 := 2)
   END_RUNG wire#w2
   RUNG wire#w1
      { S7_Templates := "SrcType := Int" } EQ_Contact(in1 := "全局数据块".手动存储仓位, in2 := 3)
   END_RUNG wire#w2
   RUNG wire#w2
      S_Coil( "运动控制数据2".X值统一入库位 )
   END_RUNG
   RUNG wire#w1
      { S7_Templates := "SrcType := Int" } EQ_Contact(in1 := "全局数据块".手动存储仓位, in2 := 4)
      wire#w3
      Move(in := "运动控制数据2".def位x值, out1 => "运动控制数据2".X轴位置)
   END_RUNG
   RUNG wire#w1
      { S7_Templates := "SrcType := Int" } EQ_Contact(in1 := "全局数据块".手动存储仓位, in2 := 5)
   END_RUNG wire#w3
   RUNG wire#w1
      { S7_Templates := "SrcType := Int" } EQ_Contact(in1 := "全局数据块".手动存储仓位, in2 := 6)
   END_RUNG wire#w3
   RUNG wire#w3
      S_Coil( "运动控制数据2".X值统一入库位 )
   END_RUNG
   RUNG wire#w1
      { S7_Templates := "SrcType := Int" } EQ_Contact(in1 := "全局数据块".手动存储仓位, in2 := 7)
      wire#w4
      Move(in := "运动控制数据2".ghi位x值, out1 => "运动控制数据2".X轴位置)
   END_RUNG
   RUNG wire#w1
      { S7_Templates := "SrcType := Int" } EQ_Contact(in1 := "全局数据块".手动存储仓位, in2 := 8)
   END_RUNG wire#w4
   RUNG wire#w1
      { S7_Templates := "SrcType := Int" } EQ_Contact(in1 := "全局数据块".手动存储仓位, in2 := 9)
   END_RUNG wire#w4
   RUNG wire#w4
      S_Coil( "运动控制数据2".X值统一入库位 )
   END_RUNG
   RUNG wire#powerrail
      { S7_Templates := "SrcType := Real" } EQ_Contact(in1 := "全局数据块".手动模式步骤, in2 := 14.0)
      wire#w5
      { S7_Templates := "SrcType := Int" } EQ_Contact(in1 := "全局数据块".手动存储仓位, in2 := 1)
      wire#w6
      Move(in := "运动控制数据2".adg位y值, out1 => "运动控制数据2".Y轴位置)
   END_RUNG
   RUNG wire#w5
      { S7_Templates := "SrcType := Int" } EQ_Contact(in1 := "全局数据块".手动存储仓位, in2 := 4)
   END_RUNG wire#w6
   RUNG wire#w5
      { S7_Templates := "SrcType := Int" } EQ_Contact(in1 := "全局数据块".手动存储仓位, in2 := 7)
   END_RUNG wire#w6
   RUNG wire#w6
      S_Coil( "运动控制数据2".Y值统一入库位 )
   END_RUNG
   RUNG wire#w5
      { S7_Templates := "SrcType := Int" } EQ_Contact(in1 := "全局数据块".手动存储仓位, in2 := 2)
      wire#w7
      Move(in := "运动控制数据2".bef位y值, out1 => "运动控制数据2".Y轴位置)
   END_RUNG
   RUNG wire#w5
      { S7_Templates := "SrcType := Int" } EQ_Contact(in1 := "全局数据块".手动存储仓位, in2 := 5)
   END_RUNG wire#w7
   RUNG wire#w5
      { S7_Templates := "SrcType := Int" } EQ_Contact(in1 := "全局数据块".手动存储仓位, in2 := 8)
   END_RUNG wire#w7
   RUNG wire#w7
      S_Coil( "运动控制数据2".Y值统一入库位 )
   END_RUNG
   RUNG wire#w5
      { S7_Templates := "SrcType := Int" } EQ_Contact(in1 := "全局数据块".手动存储仓位, in2 := 3)
      wire#w8
      Move(in := "运动控制数据2".cfi位y值, out1 => "运动控制数据2".Y轴位置)
   END_RUNG
   RUNG wire#w5
      { S7_Templates := "SrcType := Int" } EQ_Contact(in1 := "全局数据块".手动存储仓位, in2 := 6)
   END_RUNG wire#w8
   RUNG wire#w5
      { S7_Templates := "SrcType := Int" } EQ_Contact(in1 := "全局数据块".手动存储仓位, in2 := 9)
   END_RUNG wire#w8
   RUNG wire#w8
      S_Coil( "运动控制数据2".Y值统一入库位 )
   END_RUNG
   RUNG wire#powerrail
      { S7_Templates := "SrcType := Real" } EQ_Contact(in1 := "全局数据块".手动模式步骤, in2 := 14.0)
      Contact( "运动控制数据2".X值统一入库位 )
      Contact( "运动控制数据2".Y值统一入库位 )
      { S7_Templates := "SrcType := Real" } EQ_Contact(in1 := "X轴机械手".Position, in2 := "运动控制数据2".X轴位置)
      { S7_Templates := "SrcType := Real" } EQ_Contact(in1 := "Y轴机械手".Position, in2 := "运动控制数据2".Y轴位置)
      wire#w9
      Move(in := 15.0, out1 => "全局数据块".手动模式步骤)
   END_RUNG
   RUNG wire#w9
      R_Coil( "运动控制数据2".X值统一入库位 )
   END_RUNG
   RUNG wire#w9
      R_Coil( "运动控制数据2".Y值统一入库位 )
   END_RUNG
   // the same network as SCL:
   #_w1 := ("全局数据块".手动模式步骤 = 14.0) AND "[144]仓储上升位";
   IF #_w1 AND (("全局数据块".手动存储仓位 = 1) OR ("全局数据块".手动存储仓位 = 2) OR ("全局数据块".手动存储仓位 = 3)) THEN
       "运动控制数据2".X轴位置 := "运动控制数据2".abc位x值;
       "运动控制数据2".X值统一入库位 := TRUE;
   END_IF;
   IF #_w1 AND (("全局数据块".手动存储仓位 = 4) OR ("全局数据块".手动存储仓位 = 5) OR ("全局数据块".手动存储仓位 = 6)) THEN
       "运动控制数据2".X轴位置 := "运动控制数据2".def位x值;
       "运动控制数据2".X值统一入库位 := TRUE;
   END_IF;
   IF #_w1 AND (("全局数据块".手动存储仓位 = 7) OR ("全局数据块".手动存储仓位 = 8) OR ("全局数据块".手动存储仓位 = 9)) THEN
       "运动控制数据2".X轴位置 := "运动控制数据2".ghi位x值;
       "运动控制数据2".X值统一入库位 := TRUE;
   END_IF;
   #_w2 := "全局数据块".手动模式步骤 = 14.0;
   IF #_w2 AND (("全局数据块".手动存储仓位 = 1) OR ("全局数据块".手动存储仓位 = 4) OR ("全局数据块".手动存储仓位 = 7)) THEN
       "运动控制数据2".Y轴位置 := "运动控制数据2".adg位y值;
       "运动控制数据2".Y值统一入库位 := TRUE;
   END_IF;
   IF #_w2 AND (("全局数据块".手动存储仓位 = 2) OR ("全局数据块".手动存储仓位 = 5) OR ("全局数据块".手动存储仓位 = 8)) THEN
       "运动控制数据2".Y轴位置 := "运动控制数据2".bef位y值;
       "运动控制数据2".Y值统一入库位 := TRUE;
   END_IF;
   IF #_w2 AND (("全局数据块".手动存储仓位 = 3) OR ("全局数据块".手动存储仓位 = 6) OR ("全局数据块".手动存储仓位 = 9)) THEN
       "运动控制数据2".Y轴位置 := "运动控制数据2".cfi位y值;
       "运动控制数据2".Y值统一入库位 := TRUE;
   END_IF;
   #_w3 := ("全局数据块".手动模式步骤 = 14.0) AND "运动控制数据2".X值统一入库位 AND "运动控制数据2".Y值统一入库位 AND ("X轴机械手".Position = "运动控制数据2".X轴位置) AND ("Y轴机械手".Position = "运动控制数据2".Y轴位置);
   IF #_w3 THEN
       "全局数据块".手动模式步骤 := 15.0;
       "运动控制数据2".X值统一入库位 := FALSE;
       "运动控制数据2".Y值统一入库位 := FALSE;
   END_IF;
END_REGION

REGION Network 18: 放料流程
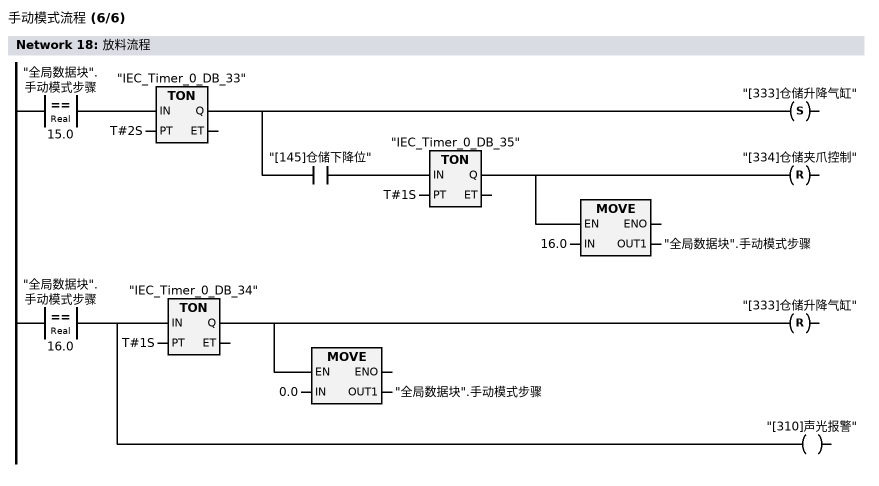
   "IEC_Timer_0_DB_33".TON(IN := "全局数据块".手动模式步骤 = 15.0, PT := T#2S);
   IF "IEC_Timer_0_DB_33".Q THEN "[333]仓储升降气缸" := TRUE; END_IF;
   "IEC_Timer_0_DB_35".TON(IN := "IEC_Timer_0_DB_33".Q AND "[145]仓储下降位", PT := T#1S);
   IF "IEC_Timer_0_DB_35".Q THEN
       "[334]仓储夹爪控制" := FALSE;
       "全局数据块".手动模式步骤 := 16.0;
   END_IF;
   #_w1 := "全局数据块".手动模式步骤 = 16.0;
   "IEC_Timer_0_DB_34".TON(IN := #_w1, PT := T#1S);
   IF "IEC_Timer_0_DB_34".Q THEN
       "[333]仓储升降气缸" := FALSE;
       "全局数据块".手动模式步骤 := 0.0;
   END_IF;
   "[310]声光报警" := #_w1;
END_REGION

REGION Network 19: 流程三入库
END_REGION
END_FUNCTION

ORGANIZATION_BLOCK "Main"   // OB1, LAD, ProgramCycle
TITLE = "Main Program Sweep (Cycle)"
{ S7_Optimized_Access := 'TRUE' }
VERSION : 0.1
   VAR_INPUT
      Initial_Call : Bool;   // Initial call of this OB
      Remanence : Bool;   // =True, if remanent data are available
   END_VAR
   VAR_TEMP   // added for the SCL form of the ladder/FBD networks
      _w1 : Bool;
      _w2 : Bool;
      _w3 : Bool;
      _w4 : Bool;
      _w5 : Bool;
      _w6 : Bool;
   END_VAR
BEGIN

REGION Network 1: 手动
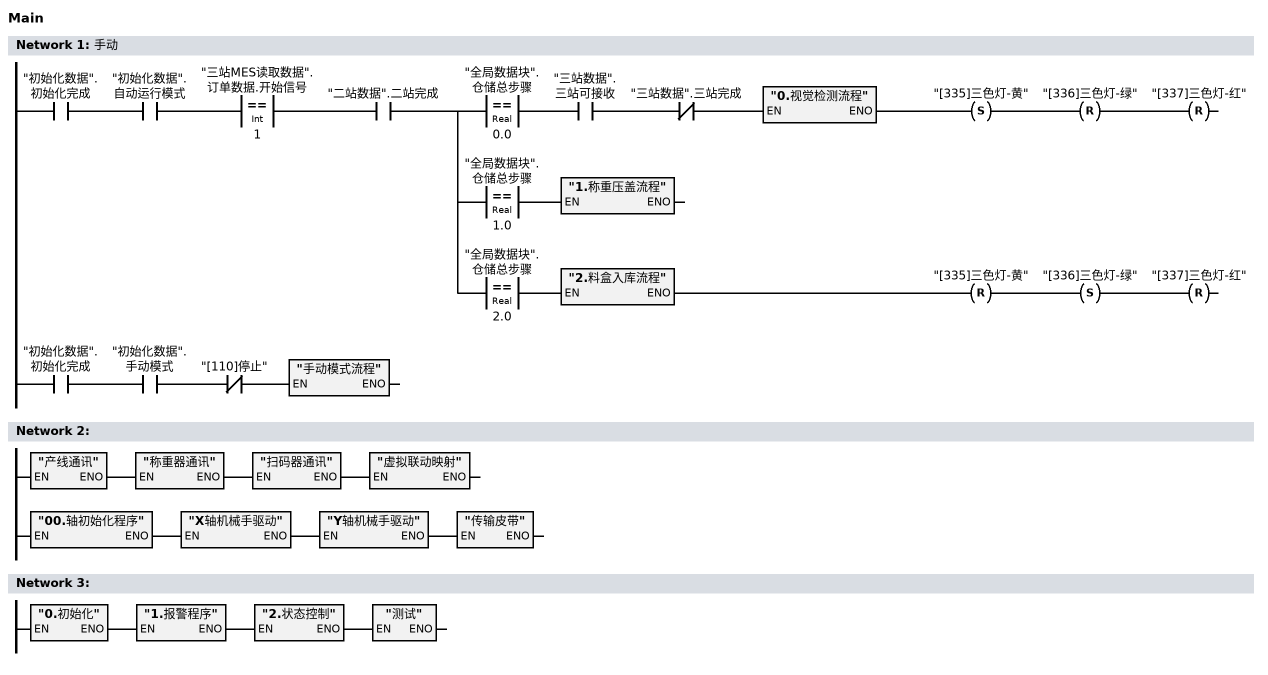
   RUNG wire#powerrail
      Contact( "初始化数据".初始化完成 )
      Contact( "初始化数据".自动运行模式 )
      { S7_Templates := "SrcType := Int" } EQ_Contact(in1 := "三站MES读取数据".订单数据.开始信号, in2 := 1)
      Contact( "二站数据".二站完成 )
      wire#w1
      { S7_Templates := "SrcType := Real" } EQ_Contact(in1 := "全局数据块".仓储总步骤, in2 := 0.0)
      Contact( "三站数据".三站可接收 )
      I_Contact( "三站数据".三站完成 )
      "0.视觉检测流程"()
      S_Coil( "[335]三色灯-黄" )
      R_Coil( "[336]三色灯-绿" )
      R_Coil( "[337]三色灯-红" )
   END_RUNG
   RUNG wire#w1
      { S7_Templates := "SrcType := Real" } EQ_Contact(in1 := "全局数据块".仓储总步骤, in2 := 1.0)
      "1.称重压盖流程"()
   END_RUNG
   RUNG wire#w1
      { S7_Templates := "SrcType := Real" } EQ_Contact(in1 := "全局数据块".仓储总步骤, in2 := 2.0)
      "2.料盒入库流程"()
      R_Coil( "[335]三色灯-黄" )
      S_Coil( "[336]三色灯-绿" )
      R_Coil( "[337]三色灯-红" )
   END_RUNG
   RUNG wire#powerrail
      Contact( "初始化数据".初始化完成 )
      Contact( "初始化数据".手动模式 )
      I_Contact( "[110]停止" )
      "手动模式流程"()
   END_RUNG
   // the same network as SCL:
   #_w1 := "初始化数据".初始化完成 AND "初始化数据".自动运行模式 AND ("三站MES读取数据".订单数据.开始信号 = 1) AND "二站数据".二站完成;
   "0.视觉检测流程"(EN := #_w1 AND ("全局数据块".仓储总步骤 = 0.0) AND "三站数据".三站可接收 AND NOT "三站数据".三站完成, ENO => #_w2);
   IF #_w2 THEN
       "[335]三色灯-黄" := TRUE;
       "[336]三色灯-绿" := FALSE;
       "[337]三色灯-红" := FALSE;
   END_IF;
   IF #_w1 AND ("全局数据块".仓储总步骤 = 1.0) THEN "1.称重压盖流程"(); END_IF;
   "2.料盒入库流程"(EN := #_w1 AND ("全局数据块".仓储总步骤 = 2.0), ENO => #_w3);
   IF #_w3 THEN
       "[335]三色灯-黄" := FALSE;
       "[336]三色灯-绿" := TRUE;
       "[337]三色灯-红" := FALSE;
   END_IF;
   IF "初始化数据".初始化完成 AND "初始化数据".手动模式 AND NOT "[110]停止" THEN "手动模式流程"(); END_IF;
END_REGION

REGION Network 2
   RUNG wire#powerrail
      "产线通讯"()
      "称重器通讯"()
      "扫码器通讯"()
      "虚拟联动映射"()
   END_RUNG
   RUNG wire#powerrail
      "00.轴初始化程序"()
      "X轴机械手驱动"()
      "Y轴机械手驱动"()
      "传输皮带"()
   END_RUNG
   // the same network as SCL:
   "产线通讯"(ENO => #_w1);
   "称重器通讯"(EN := #_w1, ENO => #_w2);
   "扫码器通讯"(EN := #_w2, ENO => #_w3);
   IF #_w3 THEN "虚拟联动映射"(); END_IF;
   "00.轴初始化程序"(ENO => #_w4);
   "X轴机械手驱动"(EN := #_w4, ENO => #_w5);
   "Y轴机械手驱动"(EN := #_w5, ENO => #_w6);
   IF #_w6 THEN "传输皮带"(); END_IF;
END_REGION

REGION Network 3
   RUNG wire#powerrail
      "0.初始化"()
      "1.报警程序"()
      "2.状态控制"()
      "测试"()
   END_RUNG
   // the same network as SCL:
   "0.初始化"(ENO => #_w1);
   "1.报警程序"(EN := #_w1, ENO => #_w2);
   "2.状态控制"(EN := #_w2, ENO => #_w3);
   IF #_w3 THEN "测试"(); END_IF;
END_REGION
END_ORGANIZATION_BLOCK

// folder: 自动模式

FUNCTION "0.视觉检测流程" : Void   // FC7, LAD
{ S7_Optimized_Access := 'TRUE' }
VERSION : 0.1
   VAR_TEMP   // added for the SCL form of the ladder/FBD networks
      _w1 : Bool;
      _w2 : Bool;
   END_VAR
BEGIN

REGION Network 1: 到拍照位
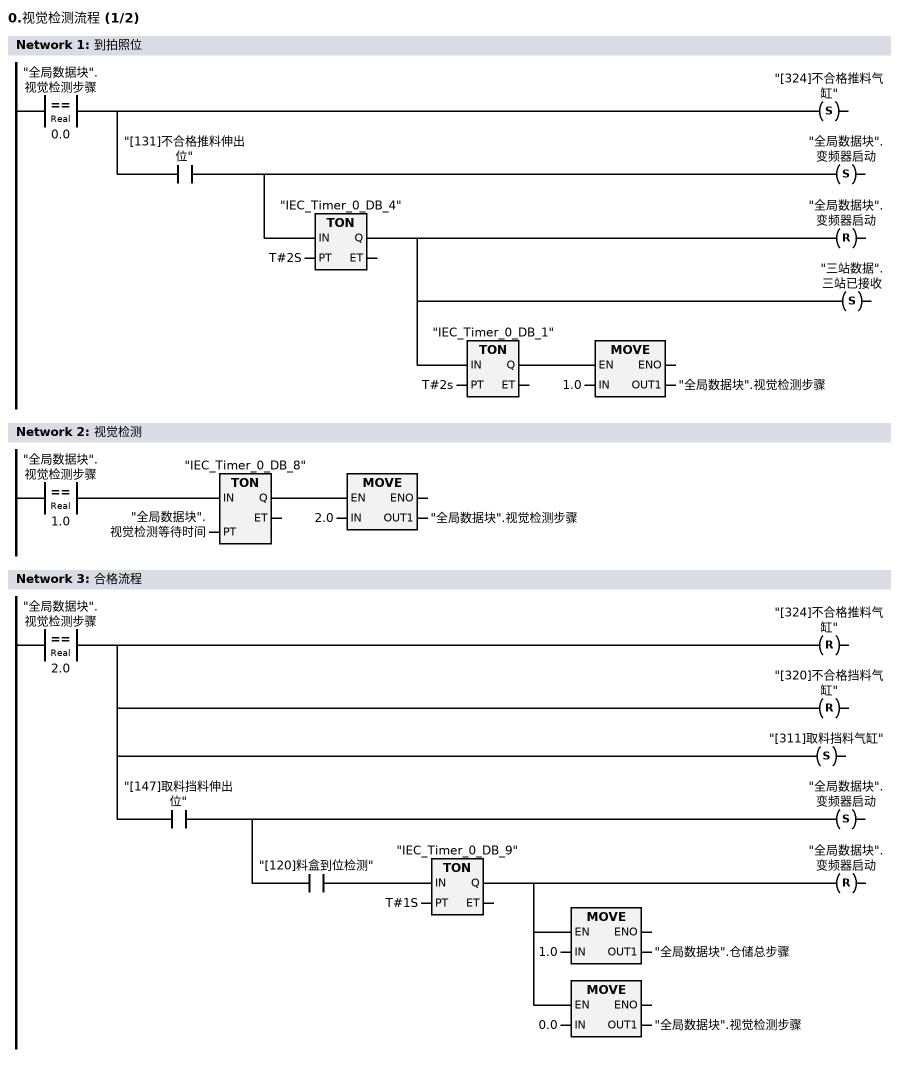
   #_w1 := "全局数据块".视觉检测步骤 = 0.0;
   IF #_w1 THEN "[324]不合格推料气缸" := TRUE; END_IF;
   #_w2 := #_w1 AND "[131]不合格推料伸出位";
   IF #_w2 THEN "全局数据块".变频器启动 := TRUE; END_IF;
   "IEC_Timer_0_DB_4".TON(IN := #_w2, PT := T#2S);
   IF "IEC_Timer_0_DB_4".Q THEN
       "全局数据块".变频器启动 := FALSE;
       "三站数据".三站已接收 := TRUE;
   END_IF;
   "IEC_Timer_0_DB_1".TON(IN := "IEC_Timer_0_DB_4".Q, PT := T#2s);
   IF "IEC_Timer_0_DB_1".Q THEN "全局数据块".视觉检测步骤 := 1.0; END_IF;
END_REGION

REGION Network 2: 视觉检测
   "IEC_Timer_0_DB_8".TON(IN := "全局数据块".视觉检测步骤 = 1.0, PT := "全局数据块".视觉检测等待时间);
   IF "IEC_Timer_0_DB_8".Q THEN "全局数据块".视觉检测步骤 := 2.0; END_IF;
END_REGION

REGION Network 3: 合格流程
   #_w1 := "全局数据块".视觉检测步骤 = 2.0;
   IF #_w1 THEN
       "[324]不合格推料气缸" := FALSE;
       "[320]不合格挡料气缸" := FALSE;
       "[311]取料挡料气缸" := TRUE;
   END_IF;
   #_w2 := #_w1 AND "[147]取料挡料伸出位";
   IF #_w2 THEN "全局数据块".变频器启动 := TRUE; END_IF;
   "IEC_Timer_0_DB_9".TON(IN := #_w2 AND "[120]料盒到位检测", PT := T#1S);
   IF "IEC_Timer_0_DB_9".Q THEN
       "全局数据块".变频器启动 := FALSE;
       "全局数据块".仓储总步骤 := 1.0;
       "全局数据块".视觉检测步骤 := 0.0;
   END_IF;
END_REGION

REGION Network 4: 不合格流程
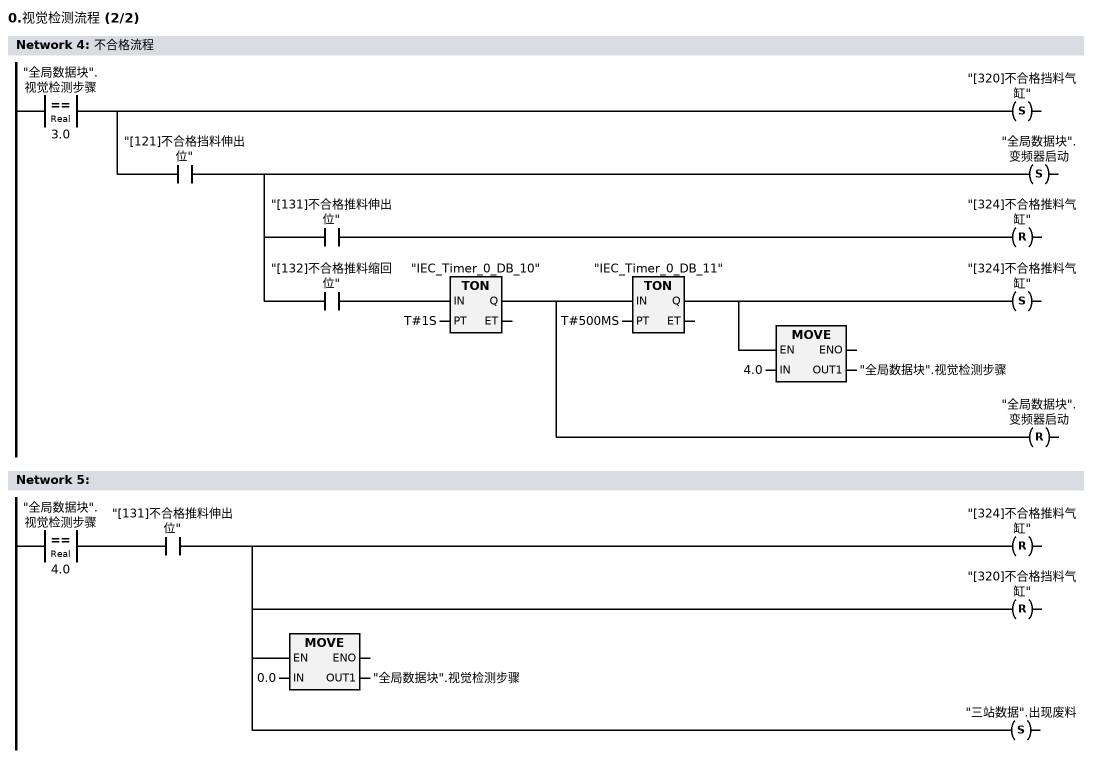
   #_w1 := "全局数据块".视觉检测步骤 = 3.0;
   IF #_w1 THEN "[320]不合格挡料气缸" := TRUE; END_IF;
   #_w2 := #_w1 AND "[121]不合格挡料伸出位";
   IF #_w2 THEN "全局数据块".变频器启动 := TRUE; END_IF;
   IF #_w2 AND "[131]不合格推料伸出位" THEN "[324]不合格推料气缸" := FALSE; END_IF;
   "IEC_Timer_0_DB_10".TON(IN := #_w2 AND "[132]不合格推料缩回位", PT := T#1S);
   "IEC_Timer_0_DB_11".TON(IN := "IEC_Timer_0_DB_10".Q, PT := T#500MS);
   IF "IEC_Timer_0_DB_11".Q THEN
       "[324]不合格推料气缸" := TRUE;
       "全局数据块".视觉检测步骤 := 4.0;
   END_IF;
   IF "IEC_Timer_0_DB_10".Q THEN "全局数据块".变频器启动 := FALSE; END_IF;
END_REGION

REGION Network 5
   RUNG wire#powerrail
      { S7_Templates := "SrcType := Real" } EQ_Contact(in1 := "全局数据块".视觉检测步骤, in2 := 4.0)
      Contact( "[131]不合格推料伸出位" )
      wire#w1
      R_Coil( "[324]不合格推料气缸" )
   END_RUNG
   RUNG wire#w1
      R_Coil( "[320]不合格挡料气缸" )
   END_RUNG
   RUNG wire#w1
      Move(in := 0.0, out1 => "全局数据块".视觉检测步骤)
   END_RUNG
   RUNG wire#w1
      S_Coil( "三站数据".出现废料 )
   END_RUNG
   // the same network as SCL:
   #_w1 := ("全局数据块".视觉检测步骤 = 4.0) AND "[131]不合格推料伸出位";
   IF #_w1 THEN
       "[324]不合格推料气缸" := FALSE;
       "[320]不合格挡料气缸" := FALSE;
       "全局数据块".视觉检测步骤 := 0.0;
       "三站数据".出现废料 := TRUE;
   END_IF;
END_REGION
END_FUNCTION

FUNCTION "1.称重压盖流程" : Void   // FC8, LAD
{ S7_Optimized_Access := 'TRUE' }
VERSION : 0.1
   VAR_TEMP   // added for the SCL form of the ladder/FBD networks
      _w1 : Bool;
      _w2 : Bool;
      _w3 : Bool;
      _w4 : Bool;
   END_VAR
BEGIN

REGION Network 1: 机械手伸出抓紧
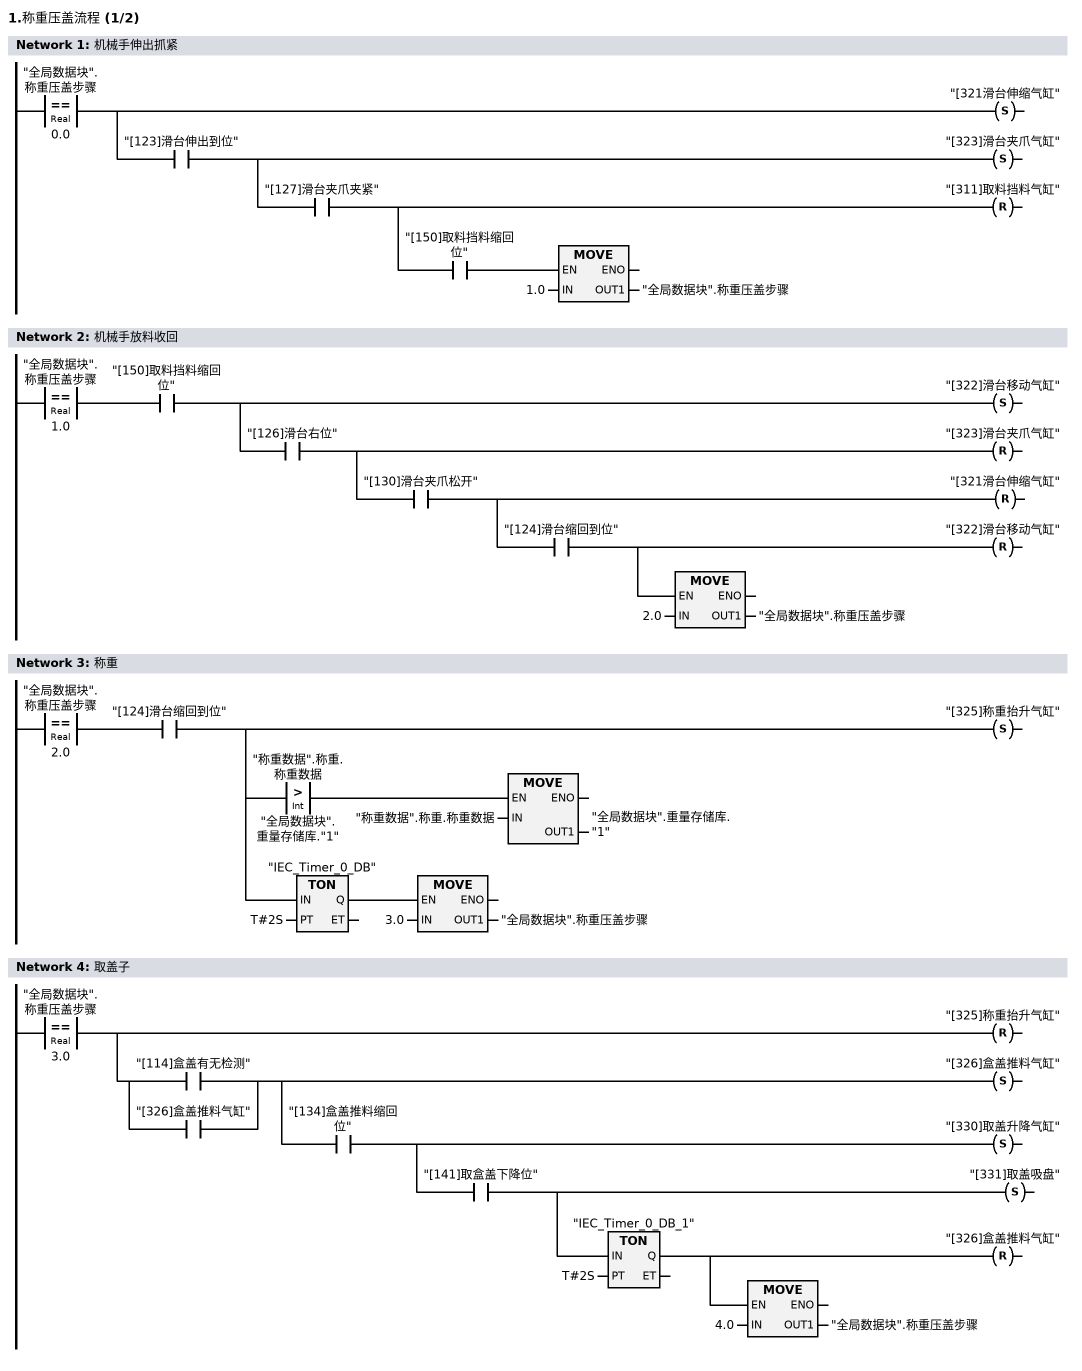
   RUNG wire#powerrail
      { S7_Templates := "SrcType := Real" } EQ_Contact(in1 := "全局数据块".称重压盖步骤, in2 := 0.0)
      wire#w1
      S_Coil( "[321滑台伸缩气缸" )
   END_RUNG
   RUNG wire#w1
      Contact( "[123]滑台伸出到位" )
      wire#w2
      S_Coil( "[323]滑台夹爪气缸" )
   END_RUNG
   RUNG wire#w2
      Contact( "[127]滑台夹爪夹紧" )
      wire#w3
      R_Coil( "[311]取料挡料气缸" )
   END_RUNG
   RUNG wire#w3
      Contact( "[150]取料挡料缩回位" )
      Move(in := 1.0, out1 => "全局数据块".称重压盖步骤)
   END_RUNG
   // the same network as SCL:
   #_w1 := "全局数据块".称重压盖步骤 = 0.0;
   IF #_w1 THEN "[321滑台伸缩气缸" := TRUE; END_IF;
   #_w2 := #_w1 AND "[123]滑台伸出到位";
   IF #_w2 THEN "[323]滑台夹爪气缸" := TRUE; END_IF;
   #_w3 := #_w2 AND "[127]滑台夹爪夹紧";
   IF #_w3 THEN "[311]取料挡料气缸" := FALSE; END_IF;
   IF #_w3 AND "[150]取料挡料缩回位" THEN "全局数据块".称重压盖步骤 := 1.0; END_IF;
END_REGION

REGION Network 2: 机械手放料收回
   RUNG wire#powerrail
      { S7_Templates := "SrcType := Real" } EQ_Contact(in1 := "全局数据块".称重压盖步骤, in2 := 1.0)
      Contact( "[150]取料挡料缩回位" )
      wire#w1
      S_Coil( "[322]滑台移动气缸" )
   END_RUNG
   RUNG wire#w1
      Contact( "[126]滑台右位" )
      wire#w2
      R_Coil( "[323]滑台夹爪气缸" )
   END_RUNG
   RUNG wire#w2
      Contact( "[130]滑台夹爪松开" )
      wire#w3
      R_Coil( "[321滑台伸缩气缸" )
   END_RUNG
   RUNG wire#w3
      Contact( "[124]滑台缩回到位" )
      wire#w4
      R_Coil( "[322]滑台移动气缸" )
   END_RUNG
   RUNG wire#w4
      Move(in := 2.0, out1 => "全局数据块".称重压盖步骤)
   END_RUNG
   // the same network as SCL:
   #_w1 := ("全局数据块".称重压盖步骤 = 1.0) AND "[150]取料挡料缩回位";
   IF #_w1 THEN "[322]滑台移动气缸" := TRUE; END_IF;
   #_w2 := #_w1 AND "[126]滑台右位";
   IF #_w2 THEN "[323]滑台夹爪气缸" := FALSE; END_IF;
   #_w3 := #_w2 AND "[130]滑台夹爪松开";
   IF #_w3 THEN "[321滑台伸缩气缸" := FALSE; END_IF;
   #_w4 := #_w3 AND "[124]滑台缩回到位";
   IF #_w4 THEN
       "[322]滑台移动气缸" := FALSE;
       "全局数据块".称重压盖步骤 := 2.0;
   END_IF;
END_REGION

REGION Network 3: 称重
   #_w1 := ("全局数据块".称重压盖步骤 = 2.0) AND "[124]滑台缩回到位";
   IF #_w1 THEN "[325]称重抬升气缸" := TRUE; END_IF;
   IF #_w1 AND ("称重数据".称重.称重数据 > "全局数据块".重量存储库."1") THEN "全局数据块".重量存储库."1" := "称重数据".称重.称重数据; END_IF;
   "IEC_Timer_0_DB".TON(IN := #_w1, PT := T#2S);
   IF "IEC_Timer_0_DB".Q THEN "全局数据块".称重压盖步骤 := 3.0; END_IF;
END_REGION

REGION Network 4: 取盖子
   #_w1 := "全局数据块".称重压盖步骤 = 3.0;
   IF #_w1 THEN "[325]称重抬升气缸" := FALSE; END_IF;
   #_w2 := #_w1 AND ("[114]盒盖有无检测" OR "[326]盒盖推料气缸");
   IF #_w2 THEN "[326]盒盖推料气缸" := TRUE; END_IF;
   #_w3 := #_w2 AND "[134]盒盖推料缩回位";
   IF #_w3 THEN "[330]取盖升降气缸" := TRUE; END_IF;
   #_w4 := #_w3 AND "[141]取盒盖下降位";
   IF #_w4 THEN "[331]取盖吸盘" := TRUE; END_IF;
   "IEC_Timer_0_DB_1".TON(IN := #_w4, PT := T#2S);
   IF "IEC_Timer_0_DB_1".Q THEN
       "[326]盒盖推料气缸" := FALSE;
       "全局数据块".称重压盖步骤 := 4.0;
   END_IF;
END_REGION

REGION Network 5: 放盖子
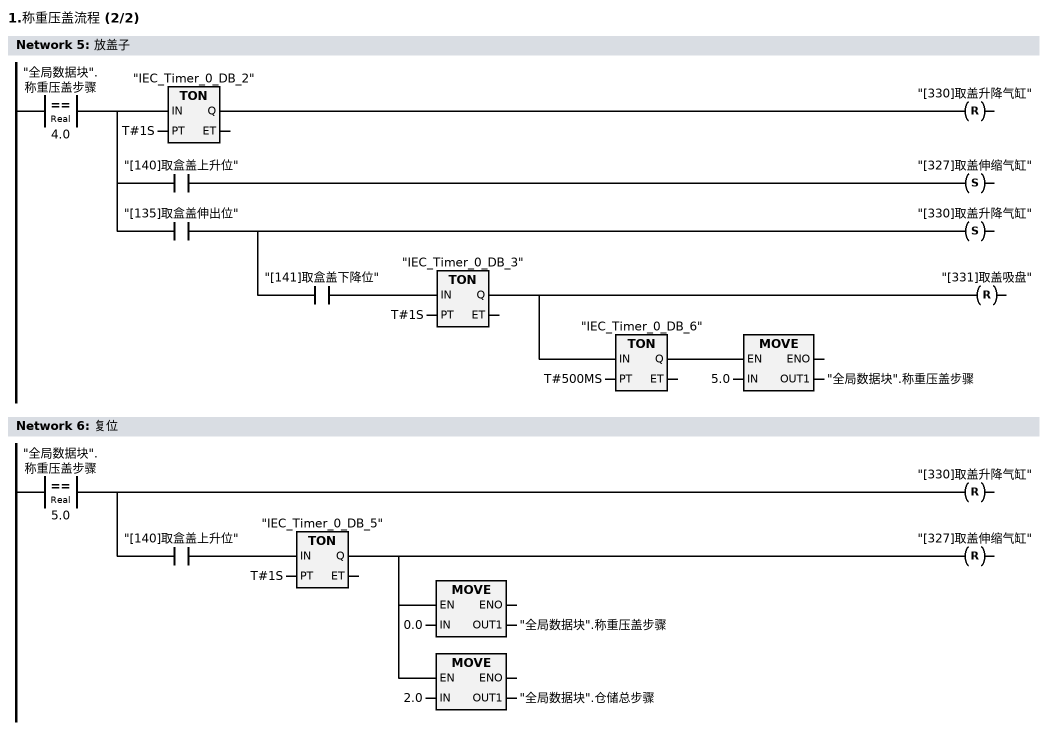
   #_w1 := "全局数据块".称重压盖步骤 = 4.0;
   "IEC_Timer_0_DB_2".TON(IN := #_w1, PT := T#1S);
   IF "IEC_Timer_0_DB_2".Q THEN "[330]取盖升降气缸" := FALSE; END_IF;
   IF #_w1 AND "[140]取盒盖上升位" THEN "[327]取盖伸缩气缸" := TRUE; END_IF;
   #_w2 := #_w1 AND "[135]取盒盖伸出位";
   IF #_w2 THEN "[330]取盖升降气缸" := TRUE; END_IF;
   "IEC_Timer_0_DB_3".TON(IN := #_w2 AND "[141]取盒盖下降位", PT := T#1S);
   IF "IEC_Timer_0_DB_3".Q THEN "[331]取盖吸盘" := FALSE; END_IF;
   "IEC_Timer_0_DB_6".TON(IN := "IEC_Timer_0_DB_3".Q, PT := T#500MS);
   IF "IEC_Timer_0_DB_6".Q THEN "全局数据块".称重压盖步骤 := 5.0; END_IF;
END_REGION

REGION Network 6: 复位
   #_w1 := "全局数据块".称重压盖步骤 = 5.0;
   IF #_w1 THEN "[330]取盖升降气缸" := FALSE; END_IF;
   "IEC_Timer_0_DB_5".TON(IN := #_w1 AND "[140]取盒盖上升位", PT := T#1S);
   IF "IEC_Timer_0_DB_5".Q THEN
       "[327]取盖伸缩气缸" := FALSE;
       "全局数据块".称重压盖步骤 := 0.0;
       "全局数据块".仓储总步骤 := 2.0;
   END_IF;
END_REGION
END_FUNCTION

FUNCTION "2.料盒入库流程" : Void   // FC9, LAD
{ S7_Optimized_Access := 'TRUE' }
VERSION : 0.1
   VAR_TEMP   // added for the SCL form of the ladder/FBD networks
      _w1 : Bool;
      _w2 : Bool;
      _w3 : Bool;
   END_VAR
BEGIN

REGION Network 1: 到取料位
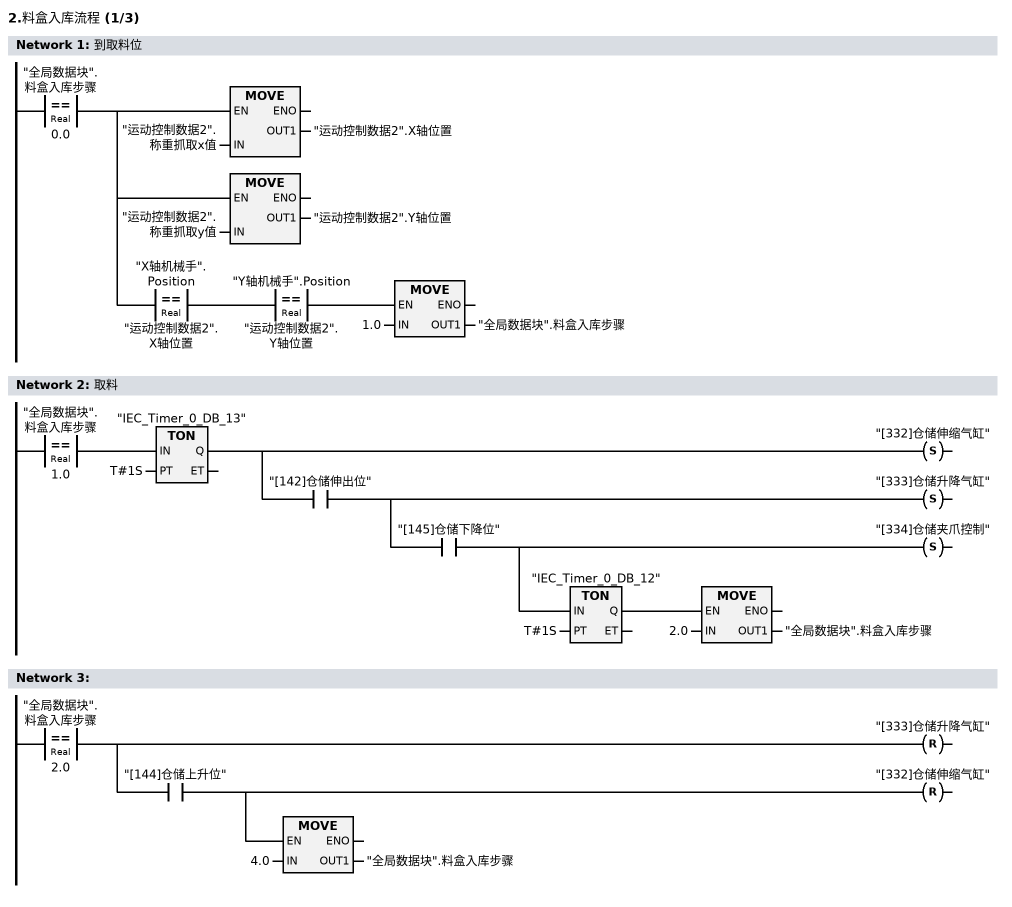
   RUNG wire#powerrail
      { S7_Templates := "SrcType := Real" } EQ_Contact(in1 := "全局数据块".料盒入库步骤, in2 := 0.0)
      wire#w1
      Move(in := "运动控制数据2".称重抓取x值, out1 => "运动控制数据2".X轴位置)
   END_RUNG
   RUNG wire#w1
      Move(in := "运动控制数据2".称重抓取y值, out1 => "运动控制数据2".Y轴位置)
   END_RUNG
   RUNG wire#w1
      { S7_Templates := "SrcType := Real" } EQ_Contact(in1 := "X轴机械手".Position, in2 := "运动控制数据2".X轴位置)
      { S7_Templates := "SrcType := Real" } EQ_Contact(in1 := "Y轴机械手".Position, in2 := "运动控制数据2".Y轴位置)
      Move(in := 1.0, out1 => "全局数据块".料盒入库步骤)
   END_RUNG
   // the same network as SCL:
   #_w1 := "全局数据块".料盒入库步骤 = 0.0;
   IF #_w1 THEN
       "运动控制数据2".X轴位置 := "运动控制数据2".称重抓取x值;
       "运动控制数据2".Y轴位置 := "运动控制数据2".称重抓取y值;
   END_IF;
   IF #_w1 AND ("X轴机械手".Position = "运动控制数据2".X轴位置) AND ("Y轴机械手".Position = "运动控制数据2".Y轴位置) THEN
       "全局数据块".料盒入库步骤 := 1.0;
   END_IF;
END_REGION

REGION Network 2: 取料
   "IEC_Timer_0_DB_13".TON(IN := "全局数据块".料盒入库步骤 = 1.0, PT := T#1S);
   IF "IEC_Timer_0_DB_13".Q THEN "[332]仓储伸缩气缸" := TRUE; END_IF;
   #_w1 := "IEC_Timer_0_DB_13".Q AND "[142]仓储伸出位";
   IF #_w1 THEN "[333]仓储升降气缸" := TRUE; END_IF;
   #_w2 := #_w1 AND "[145]仓储下降位";
   IF #_w2 THEN "[334]仓储夹爪控制" := TRUE; END_IF;
   "IEC_Timer_0_DB_12".TON(IN := #_w2, PT := T#1S);
   IF "IEC_Timer_0_DB_12".Q THEN "全局数据块".料盒入库步骤 := 2.0; END_IF;
END_REGION

REGION Network 3
   RUNG wire#powerrail
      { S7_Templates := "SrcType := Real" } EQ_Contact(in1 := "全局数据块".料盒入库步骤, in2 := 2.0)
      wire#w1
      R_Coil( "[333]仓储升降气缸" )
   END_RUNG
   RUNG wire#w1
      Contact( "[144]仓储上升位" )
      wire#w2
      R_Coil( "[332]仓储伸缩气缸" )
   END_RUNG
   RUNG wire#w2
      Move(in := 4.0, out1 => "全局数据块".料盒入库步骤)
   END_RUNG
   // the same network as SCL:
   #_w1 := "全局数据块".料盒入库步骤 = 2.0;
   IF #_w1 THEN "[333]仓储升降气缸" := FALSE; END_IF;
   #_w2 := #_w1 AND "[144]仓储上升位";
   IF #_w2 THEN
       "[332]仓储伸缩气缸" := FALSE;
       "全局数据块".料盒入库步骤 := 4.0;
   END_IF;
END_REGION

REGION Network 4: 仓位选择
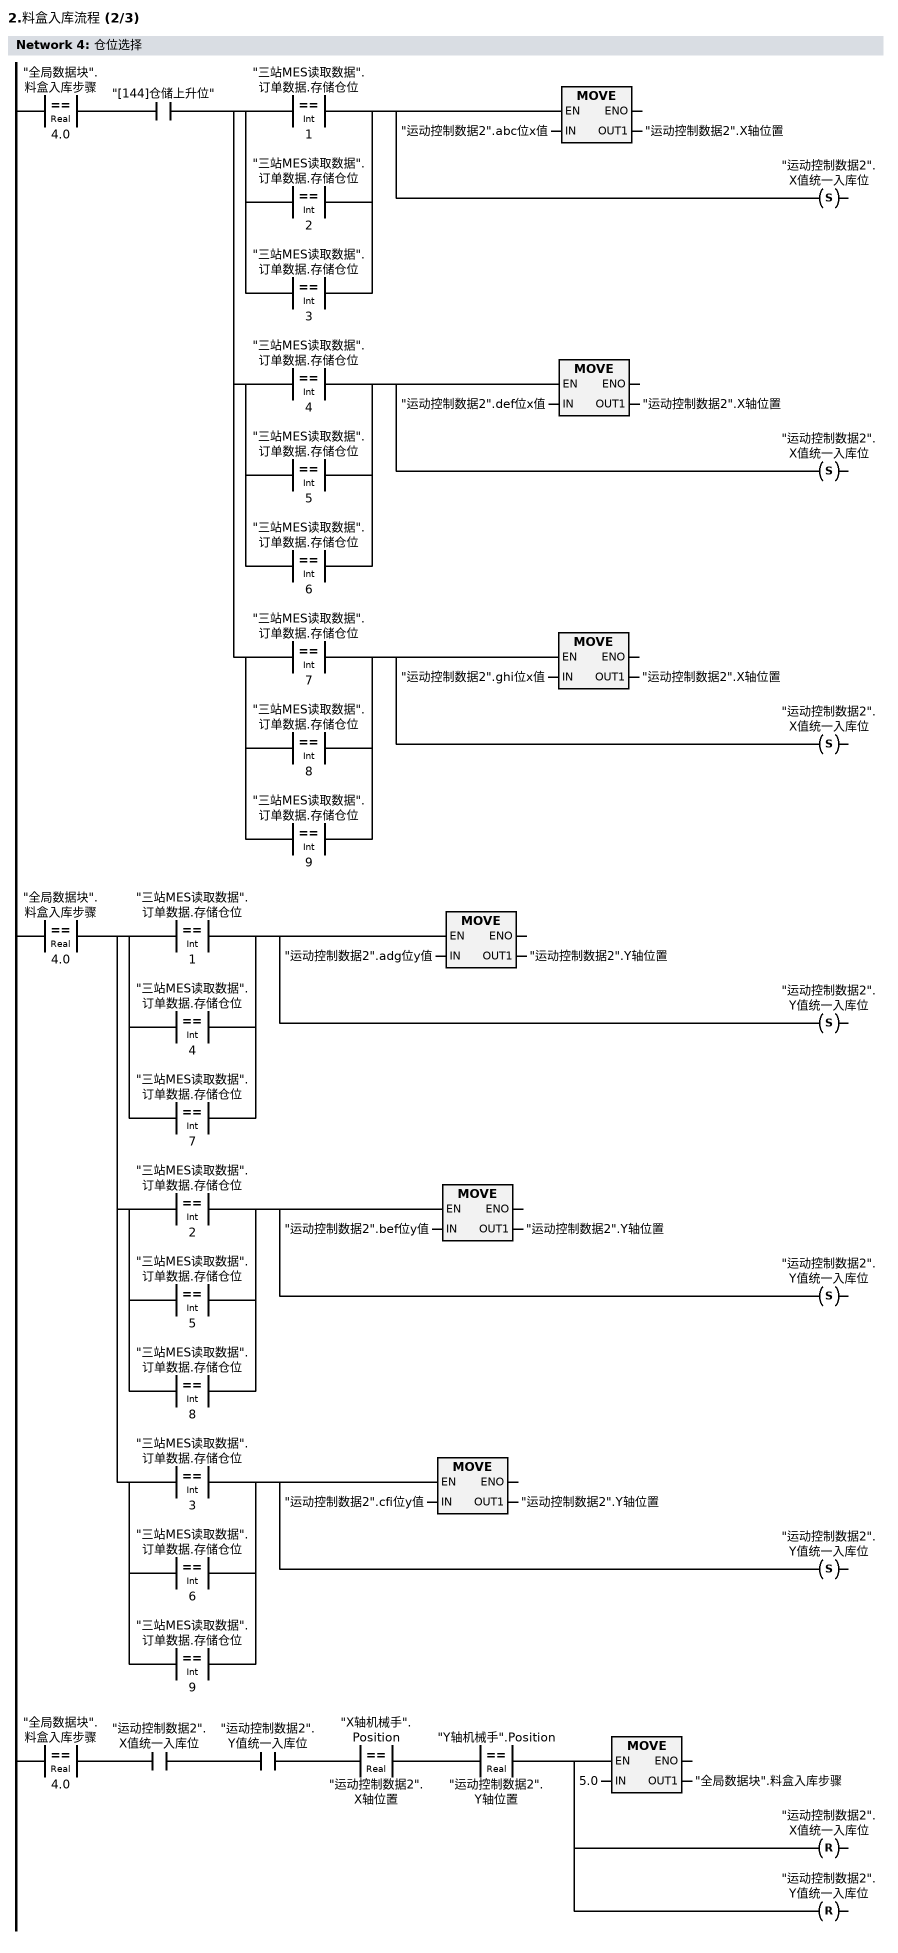
   RUNG wire#powerrail
      { S7_Templates := "SrcType := Real" } EQ_Contact(in1 := "全局数据块".料盒入库步骤, in2 := 4.0)
      Contact( "[144]仓储上升位" )
      wire#w1
      { S7_Templates := "SrcType := Int" } EQ_Contact(in1 := "三站MES读取数据".订单数据.存储仓位, in2 := 1)
      wire#w2
      Move(in := "运动控制数据2".abc位x值, out1 => "运动控制数据2".X轴位置)
   END_RUNG
   RUNG wire#w1
      { S7_Templates := "SrcType := Int" } EQ_Contact(in1 := "三站MES读取数据".订单数据.存储仓位, in2 := 2)
   END_RUNG wire#w2
   RUNG wire#w1
      { S7_Templates := "SrcType := Int" } EQ_Contact(in1 := "三站MES读取数据".订单数据.存储仓位, in2 := 3)
   END_RUNG wire#w2
   RUNG wire#w2
      S_Coil( "运动控制数据2".X值统一入库位 )
   END_RUNG
   RUNG wire#w1
      { S7_Templates := "SrcType := Int" } EQ_Contact(in1 := "三站MES读取数据".订单数据.存储仓位, in2 := 4)
      wire#w3
      Move(in := "运动控制数据2".def位x值, out1 => "运动控制数据2".X轴位置)
   END_RUNG
   RUNG wire#w1
      { S7_Templates := "SrcType := Int" } EQ_Contact(in1 := "三站MES读取数据".订单数据.存储仓位, in2 := 5)
   END_RUNG wire#w3
   RUNG wire#w1
      { S7_Templates := "SrcType := Int" } EQ_Contact(in1 := "三站MES读取数据".订单数据.存储仓位, in2 := 6)
   END_RUNG wire#w3
   RUNG wire#w3
      S_Coil( "运动控制数据2".X值统一入库位 )
   END_RUNG
   RUNG wire#w1
      { S7_Templates := "SrcType := Int" } EQ_Contact(in1 := "三站MES读取数据".订单数据.存储仓位, in2 := 7)
      wire#w4
      Move(in := "运动控制数据2".ghi位x值, out1 => "运动控制数据2".X轴位置)
   END_RUNG
   RUNG wire#w1
      { S7_Templates := "SrcType := Int" } EQ_Contact(in1 := "三站MES读取数据".订单数据.存储仓位, in2 := 8)
   END_RUNG wire#w4
   RUNG wire#w1
      { S7_Templates := "SrcType := Int" } EQ_Contact(in1 := "三站MES读取数据".订单数据.存储仓位, in2 := 9)
   END_RUNG wire#w4
   RUNG wire#w4
      S_Coil( "运动控制数据2".X值统一入库位 )
   END_RUNG
   RUNG wire#powerrail
      { S7_Templates := "SrcType := Real" } EQ_Contact(in1 := "全局数据块".料盒入库步骤, in2 := 4.0)
      wire#w5
      { S7_Templates := "SrcType := Int" } EQ_Contact(in1 := "三站MES读取数据".订单数据.存储仓位, in2 := 1)
      wire#w6
      Move(in := "运动控制数据2".adg位y值, out1 => "运动控制数据2".Y轴位置)
   END_RUNG
   RUNG wire#w5
      { S7_Templates := "SrcType := Int" } EQ_Contact(in1 := "三站MES读取数据".订单数据.存储仓位, in2 := 4)
   END_RUNG wire#w6
   RUNG wire#w5
      { S7_Templates := "SrcType := Int" } EQ_Contact(in1 := "三站MES读取数据".订单数据.存储仓位, in2 := 7)
   END_RUNG wire#w6
   RUNG wire#w6
      S_Coil( "运动控制数据2".Y值统一入库位 )
   END_RUNG
   RUNG wire#w5
      { S7_Templates := "SrcType := Int" } EQ_Contact(in1 := "三站MES读取数据".订单数据.存储仓位, in2 := 2)
      wire#w7
      Move(in := "运动控制数据2".bef位y值, out1 => "运动控制数据2".Y轴位置)
   END_RUNG
   RUNG wire#w5
      { S7_Templates := "SrcType := Int" } EQ_Contact(in1 := "三站MES读取数据".订单数据.存储仓位, in2 := 5)
   END_RUNG wire#w7
   RUNG wire#w5
      { S7_Templates := "SrcType := Int" } EQ_Contact(in1 := "三站MES读取数据".订单数据.存储仓位, in2 := 8)
   END_RUNG wire#w7
   RUNG wire#w7
      S_Coil( "运动控制数据2".Y值统一入库位 )
   END_RUNG
   RUNG wire#w5
      { S7_Templates := "SrcType := Int" } EQ_Contact(in1 := "三站MES读取数据".订单数据.存储仓位, in2 := 3)
      wire#w8
      Move(in := "运动控制数据2".cfi位y值, out1 => "运动控制数据2".Y轴位置)
   END_RUNG
   RUNG wire#w5
      { S7_Templates := "SrcType := Int" } EQ_Contact(in1 := "三站MES读取数据".订单数据.存储仓位, in2 := 6)
   END_RUNG wire#w8
   RUNG wire#w5
      { S7_Templates := "SrcType := Int" } EQ_Contact(in1 := "三站MES读取数据".订单数据.存储仓位, in2 := 9)
   END_RUNG wire#w8
   RUNG wire#w8
      S_Coil( "运动控制数据2".Y值统一入库位 )
   END_RUNG
   RUNG wire#powerrail
      { S7_Templates := "SrcType := Real" } EQ_Contact(in1 := "全局数据块".料盒入库步骤, in2 := 4.0)
      Contact( "运动控制数据2".X值统一入库位 )
      Contact( "运动控制数据2".Y值统一入库位 )
      { S7_Templates := "SrcType := Real" } EQ_Contact(in1 := "X轴机械手".Position, in2 := "运动控制数据2".X轴位置)
      { S7_Templates := "SrcType := Real" } EQ_Contact(in1 := "Y轴机械手".Position, in2 := "运动控制数据2".Y轴位置)
      wire#w9
      Move(in := 5.0, out1 => "全局数据块".料盒入库步骤)
   END_RUNG
   RUNG wire#w9
      R_Coil( "运动控制数据2".X值统一入库位 )
   END_RUNG
   RUNG wire#w9
      R_Coil( "运动控制数据2".Y值统一入库位 )
   END_RUNG
   // the same network as SCL:
   #_w1 := ("全局数据块".料盒入库步骤 = 4.0) AND "[144]仓储上升位";
   IF #_w1 AND (("三站MES读取数据".订单数据.存储仓位 = 1) OR ("三站MES读取数据".订单数据.存储仓位 = 2) OR ("三站MES读取数据".订单数据.存储仓位 = 3)) THEN
       "运动控制数据2".X轴位置 := "运动控制数据2".abc位x值;
       "运动控制数据2".X值统一入库位 := TRUE;
   END_IF;
   IF #_w1 AND (("三站MES读取数据".订单数据.存储仓位 = 4) OR ("三站MES读取数据".订单数据.存储仓位 = 5) OR ("三站MES读取数据".订单数据.存储仓位 = 6)) THEN
       "运动控制数据2".X轴位置 := "运动控制数据2".def位x值;
       "运动控制数据2".X值统一入库位 := TRUE;
   END_IF;
   IF #_w1 AND (("三站MES读取数据".订单数据.存储仓位 = 7) OR ("三站MES读取数据".订单数据.存储仓位 = 8) OR ("三站MES读取数据".订单数据.存储仓位 = 9)) THEN
       "运动控制数据2".X轴位置 := "运动控制数据2".ghi位x值;
       "运动控制数据2".X值统一入库位 := TRUE;
   END_IF;
   #_w2 := "全局数据块".料盒入库步骤 = 4.0;
   IF #_w2 AND (("三站MES读取数据".订单数据.存储仓位 = 1) OR ("三站MES读取数据".订单数据.存储仓位 = 4) OR ("三站MES读取数据".订单数据.存储仓位 = 7)) THEN
       "运动控制数据2".Y轴位置 := "运动控制数据2".adg位y值;
       "运动控制数据2".Y值统一入库位 := TRUE;
   END_IF;
   IF #_w2 AND (("三站MES读取数据".订单数据.存储仓位 = 2) OR ("三站MES读取数据".订单数据.存储仓位 = 5) OR ("三站MES读取数据".订单数据.存储仓位 = 8)) THEN
       "运动控制数据2".Y轴位置 := "运动控制数据2".bef位y值;
       "运动控制数据2".Y值统一入库位 := TRUE;
   END_IF;
   IF #_w2 AND (("三站MES读取数据".订单数据.存储仓位 = 3) OR ("三站MES读取数据".订单数据.存储仓位 = 6) OR ("三站MES读取数据".订单数据.存储仓位 = 9)) THEN
       "运动控制数据2".Y轴位置 := "运动控制数据2".cfi位y值;
       "运动控制数据2".Y值统一入库位 := TRUE;
   END_IF;
   #_w3 := ("全局数据块".料盒入库步骤 = 4.0) AND "运动控制数据2".X值统一入库位 AND "运动控制数据2".Y值统一入库位 AND ("X轴机械手".Position = "运动控制数据2".X轴位置) AND ("Y轴机械手".Position = "运动控制数据2".Y轴位置);
   IF #_w3 THEN
       "全局数据块".料盒入库步骤 := 5.0;
       "运动控制数据2".X值统一入库位 := FALSE;
       "运动控制数据2".Y值统一入库位 := FALSE;
   END_IF;
END_REGION

REGION Network 5: 放料流程
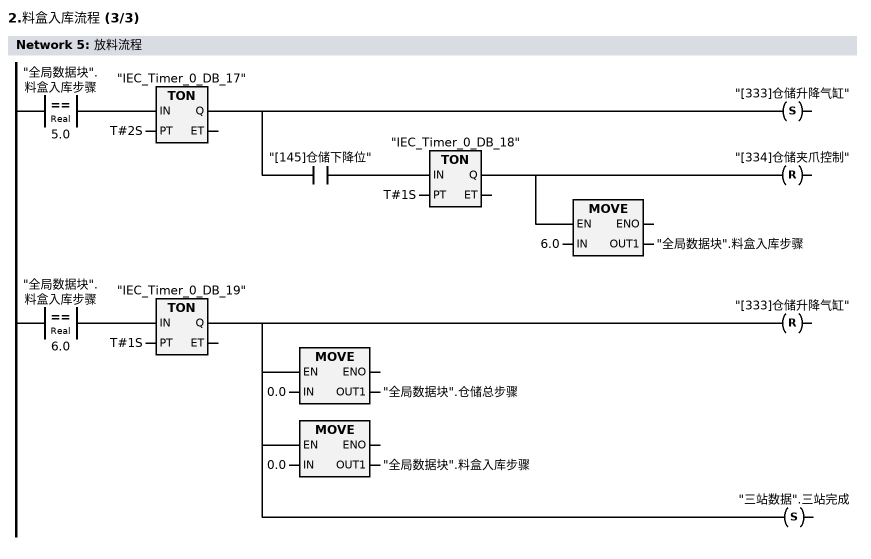
   "IEC_Timer_0_DB_17".TON(IN := "全局数据块".料盒入库步骤 = 5.0, PT := T#2S);
   IF "IEC_Timer_0_DB_17".Q THEN "[333]仓储升降气缸" := TRUE; END_IF;
   "IEC_Timer_0_DB_18".TON(IN := "IEC_Timer_0_DB_17".Q AND "[145]仓储下降位", PT := T#1S);
   IF "IEC_Timer_0_DB_18".Q THEN
       "[334]仓储夹爪控制" := FALSE;
       "全局数据块".料盒入库步骤 := 6.0;
   END_IF;
   "IEC_Timer_0_DB_19".TON(IN := "全局数据块".料盒入库步骤 = 6.0, PT := T#1S);
   IF "IEC_Timer_0_DB_19".Q THEN
       "[333]仓储升降气缸" := FALSE;
       "全局数据块".仓储总步骤 := 0.0;
       "全局数据块".料盒入库步骤 := 0.0;
       "三站数据".三站完成 := TRUE;
   END_IF;
END_REGION
END_FUNCTION

// folder: 运动控制

FUNCTION "X轴机械手驱动" : Void   // FC1, LAD
{ S7_Optimized_Access := 'TRUE' }
VERSION : 0.1
BEGIN

REGION Network 1
